PROGRAM MAIN
VAR

	fTotalCIP_Volume: REAL;
	fbWritePersistent: FB_WritePersistentData;
	bTesting		:	BOOL:=FALSE	;
	nI_1			: 	INT		;
	ftg_EStop_Fall	: 	F_TRIG	;
	rs_EStopFall	: 	RS	;
	bTestEstop		:	BOOL:=TRUE	;
	FB_OpenClose_Vlave_4026: FB_OpenClose_Vlave;
	bTemp_Water_Overweight_check: BOOL;
	fbUPS: FB_S_UPS_CX51x0;

	bSetExpeationTime: BOOL;
	i: E_ELEMENT_LIST;
	tExpirationSet_Test: TIME := T#10s;
END_VAR

prg_RealClock();
prg_Piston();
prg_Safety();
prg_MessageManager();
prg_Messages();
prg_Call_OpMode();
prg_IntCheck();
prg_User();
act_ResetPumps();
(*
prg_TriBlender(
		fb_TriBlenderPump:= g_Pump.fbPump[E_Pump_List.TB0001],
		stTriblender:=stTriblender,
		arrComponents:=arrProductionComponents);
*)		
//act_SetAnalogSens_Test();//To be deleted, for testing purposes
act_Call_Sensors_Analog();//To be deleted, for testing purposes
act_Call_Sensors_Analog_1();//To be deleted, for testing purposes
act_Call_ScaleFactor();//To be deleted, for testing purposes
act_Call_ProcessCntrl();

act_SetValves();
act_ClientPump_Select();
act_ClientStirrer_Select();
act_Call_Elements();
act_Call_Elements_Imp();
act_Call_Pumps();
prg_InterCon_Usage();
act_Sensors();
act_HeatExchenger();
act_Call_CIP();
act_Call_Production();

act_Call_For_HMI();

g_SFC.fbSFC_Temp1();

//Temtprary Overweght protection!!!!! DO NOT DELETE
IF fTotalCIP_Volume >=1500 AND FALSE THEN;
	//fbPis[E_Pis_Name.V1022].m_SetByRecipe(stPis:=stPis[E_Pis_Name.V1022], req:=E_Piston_Recipe_State.Release);
	//fbPis[E_Pis_Name.V1019].m_SetByRecipe(stPis:=stPis[E_Pis_Name.V1019], req:=E_Piston_Recipe_State.Release);
	//fbPis[E_Pis_Name.V1016].m_SetByRecipe(stPis:=stPis[E_Pis_Name.V1016], req:=E_Piston_Recipe_State.Release);
	//fbPis[E_Pis_Name.V1011].m_SetByRecipe(stPis:=stPis[E_Pis_Name.V1011], req:=E_Piston_Recipe_State.Release);
	bTemp_Water_Overweight_check:=FALSE;
	fbPrintErrMessageByID(sModuleDescription:='CIP',sActErrorID:='101x000x000');
ELSIF fTotalCIP_Volume < 1480 THEN;
	bTemp_Water_Overweight_check:=TRUE;
END_IF

IF arrTanksSens[E_Tank_Name.T91].get_stTankLevel_OverFlow() THEN;
	fbPis[E_Pis_Name.V1022].m_SetByRecipe(stPis:=stPis[E_Pis_Name.V1022], req:=E_Piston_Recipe_State.Release);
	//print error
	fbPrintErrMessageByID(sModuleDescription:='CIP',sActErrorID:='101x000x001');		
END_IF
IF arrTanksSens[E_Tank_Name.T92].get_stTankLevel_OverFlow() THEN;
	fbPis[E_Pis_Name.V1019].m_SetByRecipe(stPis:=stPis[E_Pis_Name.V1019], req:=E_Piston_Recipe_State.Release);
	//print error
	fbPrintErrMessageByID(sModuleDescription:='CIP',sActErrorID:='101x000x002');		
END_IF
IF arrTanksSens[E_Tank_Name.T93].get_stTankLevel_OverFlow() THEN;
	fbPis[E_Pis_Name.V1016].m_SetByRecipe(stPis:=stPis[E_Pis_Name.V1016], req:=E_Piston_Recipe_State.Release);
	//print error	
	fbPrintErrMessageByID(sModuleDescription:='CIP',sActErrorID:='101x000x003');	
END_IF
IF arrTanksSens[E_Tank_Name.T94].get_stTankLevel_OverFlow() THEN;
	fbPis[E_Pis_Name.V1011].m_SetByRecipe(stPis:=stPis[E_Pis_Name.V1011], req:=E_Piston_Recipe_State.Release);
	//print error
	fbPrintErrMessageByID(sModuleDescription:='CIP',sActErrorID:='101x000x004');		
END_IF
	
IF bSetExpeationTime THEN;
	bSetExpeationTime:=FALSE;
	FOR i:=E_Element_List.eTank_1 TO E_Element_List.eLine_Color DO
		fbElement[i].ExpirationTime:=tExpirationSet_Test;
		
	END_FOR
END_IF
	

mElementList_SetName();

fbWritePersistent(
	NETID:= , 
	PORT:= 851, 
	START:= , 
	TMOUT:= T#3S, 
	MODE:= , 
	BUSY=> , 
	ERR=> , 
	ERRID=> );

fbUPS();

ACTION act_Call_CIP:
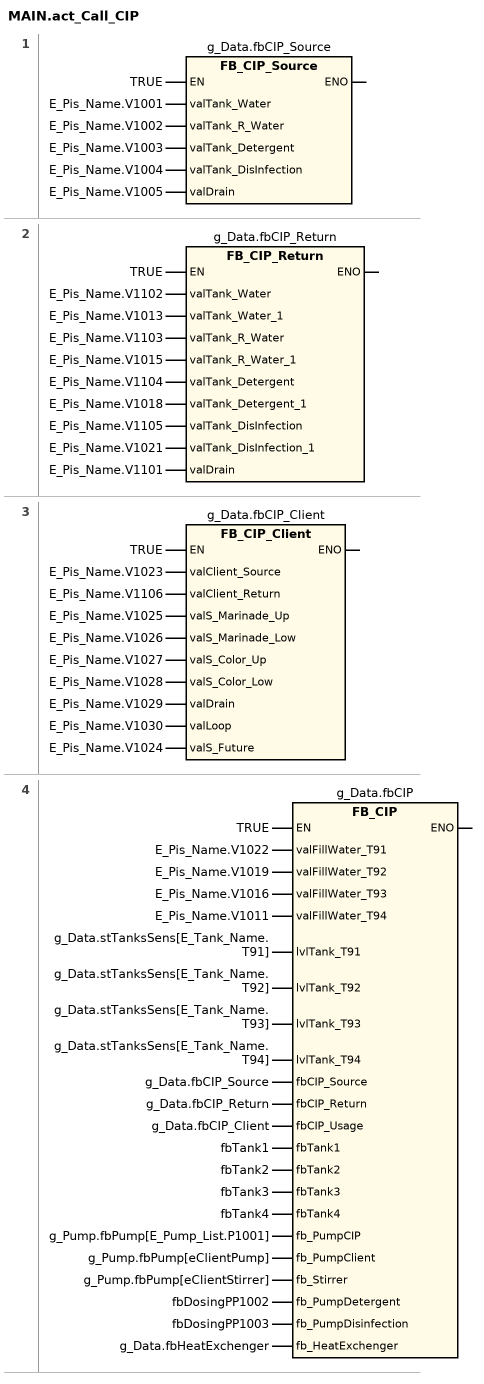
// NETWORK 1
g_Data.fbCIP_Source(
    valTank_Water := E_Pis_Name.V1001,
    valTank_R_Water := E_Pis_Name.V1002,
    valTank_Detergent := E_Pis_Name.V1003,
    valTank_DisInfection := E_Pis_Name.V1004,
    valDrain := E_Pis_Name.V1005); // FB_CIP_Source

// NETWORK 2
g_Data.fbCIP_Return(
    valTank_Water := E_Pis_Name.V1102,
    valTank_Water_1 := E_Pis_Name.V1013,
    valTank_R_Water := E_Pis_Name.V1103,
    valTank_R_Water_1 := E_Pis_Name.V1015,
    valTank_Detergent := E_Pis_Name.V1104,
    valTank_Detergent_1 := E_Pis_Name.V1018,
    valTank_DisInfection := E_Pis_Name.V1105,
    valTank_DisInfection_1 := E_Pis_Name.V1021,
    valDrain := E_Pis_Name.V1101); // FB_CIP_Return

// NETWORK 3
g_Data.fbCIP_Client(
    valClient_Source := E_Pis_Name.V1023,
    valClient_Return := E_Pis_Name.V1106,
    valS_Marinade_Up := E_Pis_Name.V1025,
    valS_Marinade_Low := E_Pis_Name.V1026,
    valS_Color_Up := E_Pis_Name.V1027,
    valS_Color_Low := E_Pis_Name.V1028,
    valDrain := E_Pis_Name.V1029,
    valLoop := E_Pis_Name.V1030,
    valS_Future := E_Pis_Name.V1024); // FB_CIP_Client

// NETWORK 4
g_Data.fbCIP(
    valFillWater_T91 := E_Pis_Name.V1022,
    valFillWater_T92 := E_Pis_Name.V1019,
    valFillWater_T93 := E_Pis_Name.V1016,
    valFillWater_T94 := E_Pis_Name.V1011,
    lvlTank_T91 := g_Data.stTanksSens[E_Tank_Name.T91],
    lvlTank_T92 := g_Data.stTanksSens[E_Tank_Name.T92],
    lvlTank_T93 := g_Data.stTanksSens[E_Tank_Name.T93],
    lvlTank_T94 := g_Data.stTanksSens[E_Tank_Name.T94],
    fbCIP_Source := g_Data.fbCIP_Source,
    fbCIP_Return := g_Data.fbCIP_Return,
    fbCIP_Usage := g_Data.fbCIP_Client,
    fbTank1 := fbTank1,
    fbTank2 := fbTank2,
    fbTank3 := fbTank3,
    fbTank4 := fbTank4,
    fb_PumpCIP := g_Pump.fbPump[E_Pump_List.P1001],
    fb_PumpClient := g_Pump.fbPump[eClientPump],
    fb_Stirrer := g_Pump.fbPump[eClientStirrer],
    fb_PumpDetergent := fbDosingPP1002,
    fb_PumpDisinfection := fbDosingPP1003,
    fb_HeatExchenger := g_Data.fbHeatExchenger); // FB_CIP

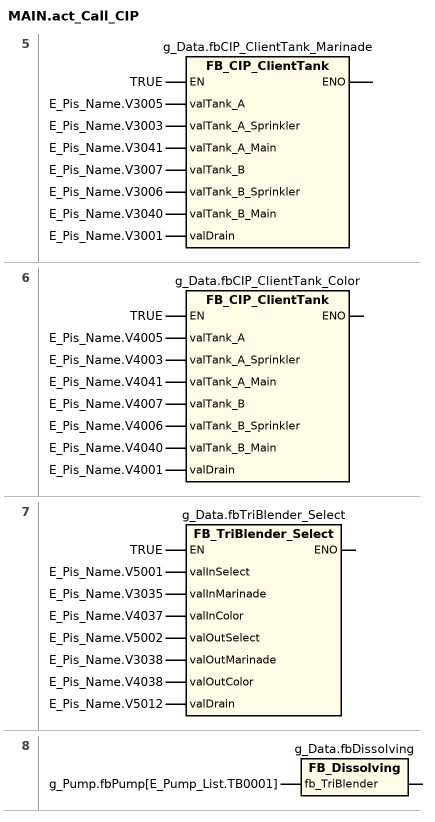
// NETWORK 5
g_Data.fbCIP_ClientTank_Marinade(
    valTank_A := E_Pis_Name.V3005,
    valTank_A_Sprinkler := E_Pis_Name.V3003,
    valTank_A_Main := E_Pis_Name.V3041,
    valTank_B := E_Pis_Name.V3007,
    valTank_B_Sprinkler := E_Pis_Name.V3006,
    valTank_B_Main := E_Pis_Name.V3040,
    valDrain := E_Pis_Name.V3001); // FB_CIP_ClientTank

// NETWORK 6
g_Data.fbCIP_ClientTank_Color(
    valTank_A := E_Pis_Name.V4005,
    valTank_A_Sprinkler := E_Pis_Name.V4003,
    valTank_A_Main := E_Pis_Name.V4041,
    valTank_B := E_Pis_Name.V4007,
    valTank_B_Sprinkler := E_Pis_Name.V4006,
    valTank_B_Main := E_Pis_Name.V4040,
    valDrain := E_Pis_Name.V4001); // FB_CIP_ClientTank

// NETWORK 7
g_Data.fbTriBlender_Select(
    valInSelect := E_Pis_Name.V5001,
    valInMarinade := E_Pis_Name.V3035,
    valInColor := E_Pis_Name.V4037,
    valOutSelect := E_Pis_Name.V5002,
    valOutMarinade := E_Pis_Name.V3038,
    valOutColor := E_Pis_Name.V4038,
    valDrain := E_Pis_Name.V5012); // FB_TriBlender_Select

// NETWORK 8
g_Data.fbDissolving(fb_TriBlender := g_Pump.fbPump[E_Pump_List.TB0001]); // FB_Dissolving
END_ACTION

ACTION act_Call_Elements:
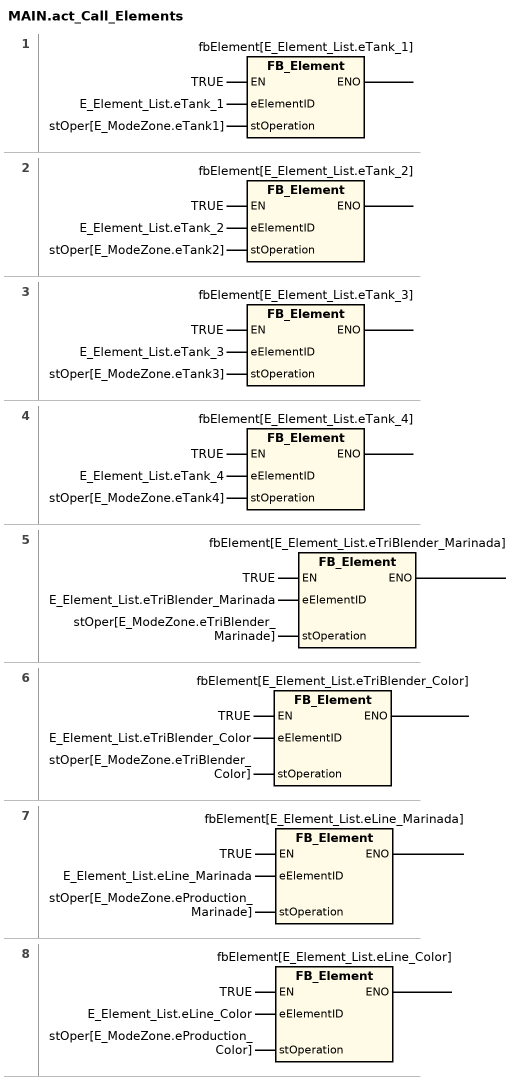
// NETWORK 1
fbElement[E_Element_List.eTank_1](eElementID := E_Element_List.eTank_1, stOperation := stOper[E_ModeZone.eTank1]); // FB_Element

// NETWORK 2
fbElement[E_Element_List.eTank_2](eElementID := E_Element_List.eTank_2, stOperation := stOper[E_ModeZone.eTank2]); // FB_Element

// NETWORK 3
fbElement[E_Element_List.eTank_3](eElementID := E_Element_List.eTank_3, stOperation := stOper[E_ModeZone.eTank3]); // FB_Element

// NETWORK 4
fbElement[E_Element_List.eTank_4](eElementID := E_Element_List.eTank_4, stOperation := stOper[E_ModeZone.eTank4]); // FB_Element

// NETWORK 5
fbElement[E_Element_List.eTriBlender_Marinada](eElementID := E_Element_List.eTriBlender_Marinada, stOperation := stOper[E_ModeZone.eTriBlender_Marinade]); // FB_Element

// NETWORK 6
fbElement[E_Element_List.eTriBlender_Color](eElementID := E_Element_List.eTriBlender_Color, stOperation := stOper[E_ModeZone.eTriBlender_Color]); // FB_Element

// NETWORK 7
fbElement[E_Element_List.eLine_Marinada](eElementID := E_Element_List.eLine_Marinada, stOperation := stOper[E_ModeZone.eProduction_Marinade]); // FB_Element

// NETWORK 8
fbElement[E_Element_List.eLine_Color](eElementID := E_Element_List.eLine_Color, stOperation := stOper[E_ModeZone.eProduction_Color]); // FB_Element
END_ACTION

ACTION act_Call_Elements_Imp:
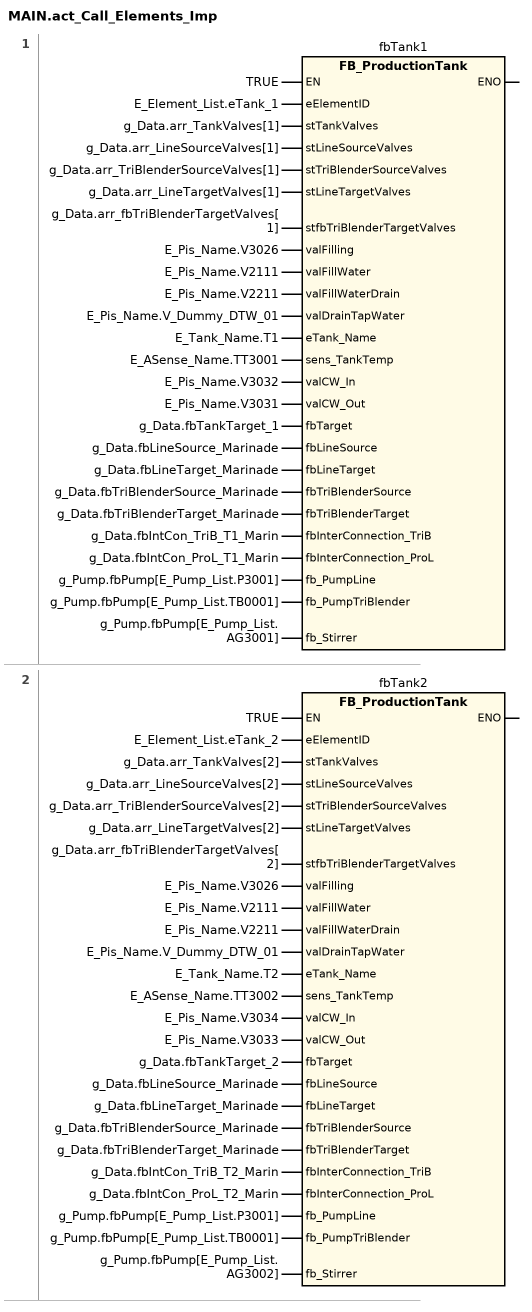
// NETWORK 1
fbTank1(
    eElementID := E_Element_List.eTank_1,
    stTankValves := g_Data.arr_TankValves[1],
    stLineSourceValves := g_Data.arr_LineSourceValves[1],
    stTriBlenderSourceValves := g_Data.arr_TriBlenderSourceValves[1],
    stLineTargetValves := g_Data.arr_LineTargetValves[1],
    stfbTriBlenderTargetValves := g_Data.arr_fbTriBlenderTargetValves[1],
    valFilling := E_Pis_Name.V3026,
    valFillWater := E_Pis_Name.V2111,
    valFillWaterDrain := E_Pis_Name.V2211,
    valDrainTapWater := E_Pis_Name.V_Dummy_DTW_01,
    eTank_Name := E_Tank_Name.T1,
    sens_TankTemp := E_ASense_Name.TT3001,
    valCW_In := E_Pis_Name.V3032,
    valCW_Out := E_Pis_Name.V3031,
    fbTarget := g_Data.fbTankTarget_1,
    fbLineSource := g_Data.fbLineSource_Marinade,
    fbLineTarget := g_Data.fbLineTarget_Marinade,
    fbTriBlenderSource := g_Data.fbTriBlenderSource_Marinade,
    fbTriBlenderTarget := g_Data.fbTriBlenderTarget_Marinade,
    fbInterConnection_TriB := g_Data.fbIntCon_TriB_T1_Marin,
    fbInterConnection_ProL := g_Data.fbIntCon_ProL_T1_Marin,
    fb_PumpLine := g_Pump.fbPump[E_Pump_List.P3001],
    fb_PumpTriBlender := g_Pump.fbPump[E_Pump_List.TB0001],
    fb_Stirrer := g_Pump.fbPump[E_Pump_List.AG3001]); // FB_ProductionTank

// NETWORK 2
fbTank2(
    eElementID := E_Element_List.eTank_2,
    stTankValves := g_Data.arr_TankValves[2],
    stLineSourceValves := g_Data.arr_LineSourceValves[2],
    stTriBlenderSourceValves := g_Data.arr_TriBlenderSourceValves[2],
    stLineTargetValves := g_Data.arr_LineTargetValves[2],
    stfbTriBlenderTargetValves := g_Data.arr_fbTriBlenderTargetValves[2],
    valFilling := E_Pis_Name.V3026,
    valFillWater := E_Pis_Name.V2111,
    valFillWaterDrain := E_Pis_Name.V2211,
    valDrainTapWater := E_Pis_Name.V_Dummy_DTW_01,
    eTank_Name := E_Tank_Name.T2,
    sens_TankTemp := E_ASense_Name.TT3002,
    valCW_In := E_Pis_Name.V3034,
    valCW_Out := E_Pis_Name.V3033,
    fbTarget := g_Data.fbTankTarget_2,
    fbLineSource := g_Data.fbLineSource_Marinade,
    fbLineTarget := g_Data.fbLineTarget_Marinade,
    fbTriBlenderSource := g_Data.fbTriBlenderSource_Marinade,
    fbTriBlenderTarget := g_Data.fbTriBlenderTarget_Marinade,
    fbInterConnection_TriB := g_Data.fbIntCon_TriB_T2_Marin,
    fbInterConnection_ProL := g_Data.fbIntCon_ProL_T2_Marin,
    fb_PumpLine := g_Pump.fbPump[E_Pump_List.P3001],
    fb_PumpTriBlender := g_Pump.fbPump[E_Pump_List.TB0001],
    fb_Stirrer := g_Pump.fbPump[E_Pump_List.AG3002]); // FB_ProductionTank

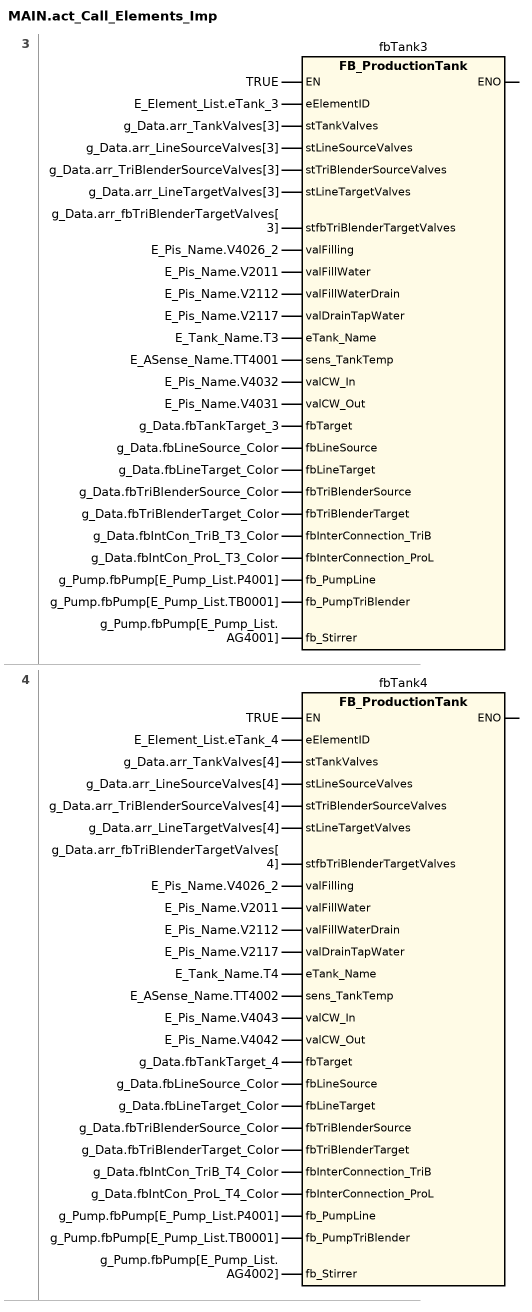
// NETWORK 3
fbTank3(
    eElementID := E_Element_List.eTank_3,
    stTankValves := g_Data.arr_TankValves[3],
    stLineSourceValves := g_Data.arr_LineSourceValves[3],
    stTriBlenderSourceValves := g_Data.arr_TriBlenderSourceValves[3],
    stLineTargetValves := g_Data.arr_LineTargetValves[3],
    stfbTriBlenderTargetValves := g_Data.arr_fbTriBlenderTargetValves[3],
    valFilling := E_Pis_Name.V4026_2,
    valFillWater := E_Pis_Name.V2011,
    valFillWaterDrain := E_Pis_Name.V2112,
    valDrainTapWater := E_Pis_Name.V2117,
    eTank_Name := E_Tank_Name.T3,
    sens_TankTemp := E_ASense_Name.TT4001,
    valCW_In := E_Pis_Name.V4032,
    valCW_Out := E_Pis_Name.V4031,
    fbTarget := g_Data.fbTankTarget_3,
    fbLineSource := g_Data.fbLineSource_Color,
    fbLineTarget := g_Data.fbLineTarget_Color,
    fbTriBlenderSource := g_Data.fbTriBlenderSource_Color,
    fbTriBlenderTarget := g_Data.fbTriBlenderTarget_Color,
    fbInterConnection_TriB := g_Data.fbIntCon_TriB_T3_Color,
    fbInterConnection_ProL := g_Data.fbIntCon_ProL_T3_Color,
    fb_PumpLine := g_Pump.fbPump[E_Pump_List.P4001],
    fb_PumpTriBlender := g_Pump.fbPump[E_Pump_List.TB0001],
    fb_Stirrer := g_Pump.fbPump[E_Pump_List.AG4001]); // FB_ProductionTank

// NETWORK 4
fbTank4(
    eElementID := E_Element_List.eTank_4,
    stTankValves := g_Data.arr_TankValves[4],
    stLineSourceValves := g_Data.arr_LineSourceValves[4],
    stTriBlenderSourceValves := g_Data.arr_TriBlenderSourceValves[4],
    stLineTargetValves := g_Data.arr_LineTargetValves[4],
    stfbTriBlenderTargetValves := g_Data.arr_fbTriBlenderTargetValves[4],
    valFilling := E_Pis_Name.V4026_2,
    valFillWater := E_Pis_Name.V2011,
    valFillWaterDrain := E_Pis_Name.V2112,
    valDrainTapWater := E_Pis_Name.V2117,
    eTank_Name := E_Tank_Name.T4,
    sens_TankTemp := E_ASense_Name.TT4002,
    valCW_In := E_Pis_Name.V4043,
    valCW_Out := E_Pis_Name.V4042,
    fbTarget := g_Data.fbTankTarget_4,
    fbLineSource := g_Data.fbLineSource_Color,
    fbLineTarget := g_Data.fbLineTarget_Color,
    fbTriBlenderSource := g_Data.fbTriBlenderSource_Color,
    fbTriBlenderTarget := g_Data.fbTriBlenderTarget_Color,
    fbInterConnection_TriB := g_Data.fbIntCon_TriB_T4_Color,
    fbInterConnection_ProL := g_Data.fbIntCon_ProL_T4_Color,
    fb_PumpLine := g_Pump.fbPump[E_Pump_List.P4001],
    fb_PumpTriBlender := g_Pump.fbPump[E_Pump_List.TB0001],
    fb_Stirrer := g_Pump.fbPump[E_Pump_List.AG4002]); // FB_ProductionTank
END_ACTION

ACTION act_Call_For_HMI:


g_HMI.stT91_Sens:=g_Data.stTanksSens[E_Tank_Name.T91];
g_HMI.stT92_Sens:=g_Data.stTanksSens[E_Tank_Name.T92];
g_HMI.stT93_Sens:=g_Data.stTanksSens[E_Tank_Name.T93];
g_HMI.stT94_Sens:=g_Data.stTanksSens[E_Tank_Name.T94];

g_HMI.stT1_Sens:=g_Data.stTanksSens[E_Tank_Name.T1];
g_HMI.stT2_Sens:=g_Data.stTanksSens[E_Tank_Name.T2];
g_HMI.stT3_Sens:=g_Data.stTanksSens[E_Tank_Name.T3];
g_HMI.stT4_Sens:=g_Data.stTanksSens[E_Tank_Name.T4];
END_ACTION

ACTION act_Call_ProcessCntrl:
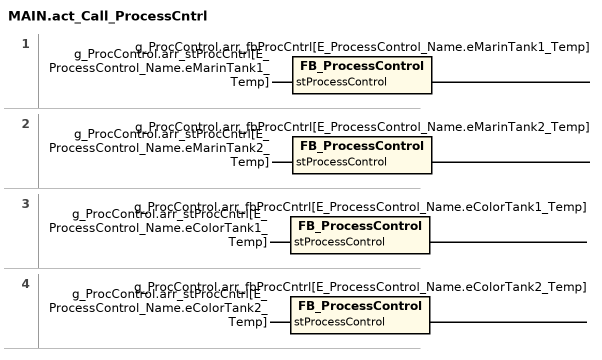
// NETWORK 1
g_ProcControl.arr_fbProcCntrl[E_ProcessControl_Name.eMarinTank1_Temp](stProcessControl := g_ProcControl.arr_stProcCntrl[E_ProcessControl_Name.eMarinTank1_Temp]); // FB_ProcessControl

// NETWORK 2
g_ProcControl.arr_fbProcCntrl[E_ProcessControl_Name.eMarinTank2_Temp](stProcessControl := g_ProcControl.arr_stProcCntrl[E_ProcessControl_Name.eMarinTank2_Temp]); // FB_ProcessControl

// NETWORK 3
g_ProcControl.arr_fbProcCntrl[E_ProcessControl_Name.eColorTank1_Temp](stProcessControl := g_ProcControl.arr_stProcCntrl[E_ProcessControl_Name.eColorTank1_Temp]); // FB_ProcessControl

// NETWORK 4
g_ProcControl.arr_fbProcCntrl[E_ProcessControl_Name.eColorTank2_Temp](stProcessControl := g_ProcControl.arr_stProcCntrl[E_ProcessControl_Name.eColorTank2_Temp]); // FB_ProcessControl
END_ACTION

ACTION act_Call_Production:

g_Prod.fbProdRecipe_Manage();
END_ACTION

ACTION act_Call_Pump_TB:
IF fbElement[E_Element_List.eTriBlender_Color].m_Get_InterConnection()=E_InterConnection.ConnToCIP 
OR fbElement[E_Element_List.eTriBlender_Marinada].m_Get_InterConnection()=E_InterConnection.ConnToCIP 
OR FALSE
THEN;
	act_Call_Pump_TB_CIP();
ELSE;
	CASE g_Data.eTriBlenderUsage OF
		E_TriBlenderUsage.eMarinada_T1,E_TriBlenderUsage.eMarinada_T2:;
				act_Call_Pump_TB_M();
		E_TriBlenderUsage.eColor_T3,E_TriBlenderUsage.eColor_T4:;
				act_Call_Pump_TB_C();
	ELSE;
		act_Call_Pump_TB_0();
	END_CASE	
END_IF
END_ACTION

ACTION act_Call_Pump_TB_0:
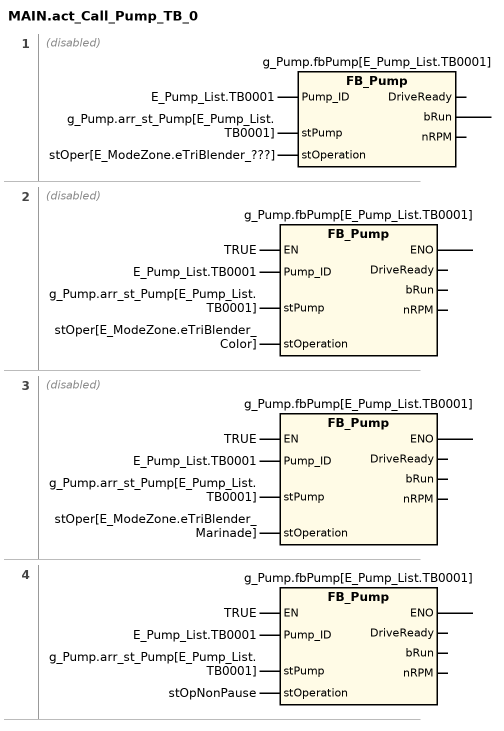
// NETWORK 1 (disabled)
// g_Pump.fbPump[E_Pump_List.TB0001](
//     Pump_ID := E_Pump_List.TB0001,
//     stPump := g_Pump.arr_st_Pump[E_Pump_List.TB0001],
//     stOperation := stOper[E_ModeZone.eTriBlender_???]); // FB_Pump

// NETWORK 2 (disabled)
// g_Pump.fbPump[E_Pump_List.TB0001](
//     Pump_ID := E_Pump_List.TB0001,
//     stPump := g_Pump.arr_st_Pump[E_Pump_List.TB0001],
//     stOperation := stOper[E_ModeZone.eTriBlender_Color]); // FB_Pump

// NETWORK 3 (disabled)
// g_Pump.fbPump[E_Pump_List.TB0001](
//     Pump_ID := E_Pump_List.TB0001,
//     stPump := g_Pump.arr_st_Pump[E_Pump_List.TB0001],
//     stOperation := stOper[E_ModeZone.eTriBlender_Marinade]); // FB_Pump

// NETWORK 4
g_Pump.fbPump[E_Pump_List.TB0001](
    Pump_ID := E_Pump_List.TB0001,
    stPump := g_Pump.arr_st_Pump[E_Pump_List.TB0001],
    stOperation := stOpNonPause); // FB_Pump
END_ACTION

ACTION act_Call_Pump_TB_C:
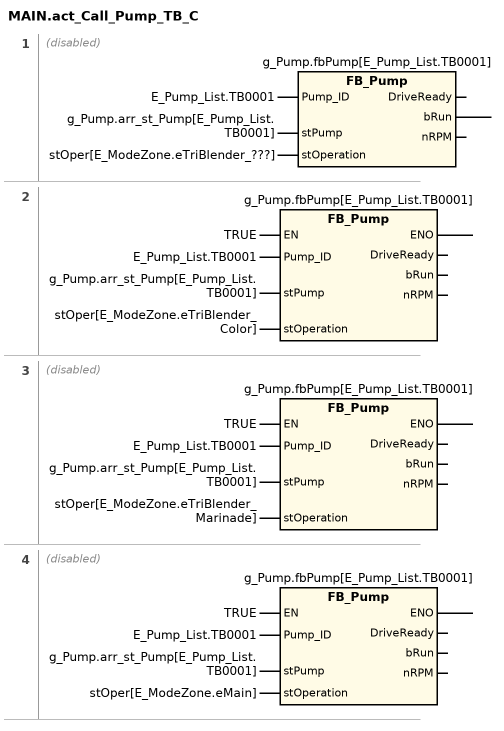
// NETWORK 1 (disabled)
// g_Pump.fbPump[E_Pump_List.TB0001](
//     Pump_ID := E_Pump_List.TB0001,
//     stPump := g_Pump.arr_st_Pump[E_Pump_List.TB0001],
//     stOperation := stOper[E_ModeZone.eTriBlender_???]); // FB_Pump

// NETWORK 2
g_Pump.fbPump[E_Pump_List.TB0001](
    Pump_ID := E_Pump_List.TB0001,
    stPump := g_Pump.arr_st_Pump[E_Pump_List.TB0001],
    stOperation := stOper[E_ModeZone.eTriBlender_Color]); // FB_Pump

// NETWORK 3 (disabled)
// g_Pump.fbPump[E_Pump_List.TB0001](
//     Pump_ID := E_Pump_List.TB0001,
//     stPump := g_Pump.arr_st_Pump[E_Pump_List.TB0001],
//     stOperation := stOper[E_ModeZone.eTriBlender_Marinade]); // FB_Pump

// NETWORK 4 (disabled)
// g_Pump.fbPump[E_Pump_List.TB0001](
//     Pump_ID := E_Pump_List.TB0001,
//     stPump := g_Pump.arr_st_Pump[E_Pump_List.TB0001],
//     stOperation := stOper[E_ModeZone.eMain]); // FB_Pump
END_ACTION

ACTION act_Call_Pump_TB_CIP:
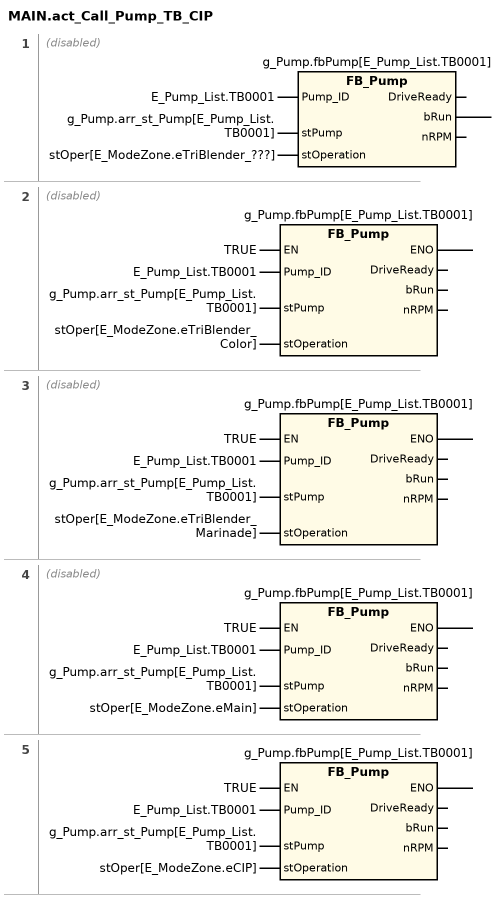
// NETWORK 1 (disabled)
// g_Pump.fbPump[E_Pump_List.TB0001](
//     Pump_ID := E_Pump_List.TB0001,
//     stPump := g_Pump.arr_st_Pump[E_Pump_List.TB0001],
//     stOperation := stOper[E_ModeZone.eTriBlender_???]); // FB_Pump

// NETWORK 2 (disabled)
// g_Pump.fbPump[E_Pump_List.TB0001](
//     Pump_ID := E_Pump_List.TB0001,
//     stPump := g_Pump.arr_st_Pump[E_Pump_List.TB0001],
//     stOperation := stOper[E_ModeZone.eTriBlender_Color]); // FB_Pump

// NETWORK 3 (disabled)
// g_Pump.fbPump[E_Pump_List.TB0001](
//     Pump_ID := E_Pump_List.TB0001,
//     stPump := g_Pump.arr_st_Pump[E_Pump_List.TB0001],
//     stOperation := stOper[E_ModeZone.eTriBlender_Marinade]); // FB_Pump

// NETWORK 4 (disabled)
// g_Pump.fbPump[E_Pump_List.TB0001](
//     Pump_ID := E_Pump_List.TB0001,
//     stPump := g_Pump.arr_st_Pump[E_Pump_List.TB0001],
//     stOperation := stOper[E_ModeZone.eMain]); // FB_Pump

// NETWORK 5
g_Pump.fbPump[E_Pump_List.TB0001](
    Pump_ID := E_Pump_List.TB0001,
    stPump := g_Pump.arr_st_Pump[E_Pump_List.TB0001],
    stOperation := stOper[E_ModeZone.eCIP]); // FB_Pump
END_ACTION

ACTION act_Call_Pump_TB_M:
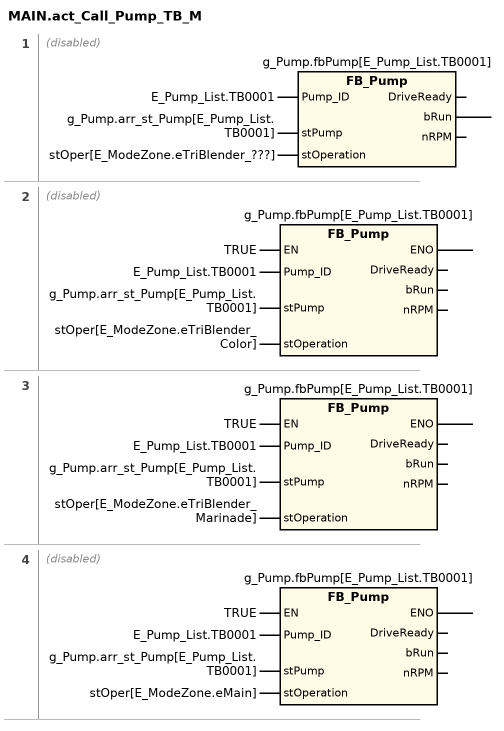
// NETWORK 1 (disabled)
// g_Pump.fbPump[E_Pump_List.TB0001](
//     Pump_ID := E_Pump_List.TB0001,
//     stPump := g_Pump.arr_st_Pump[E_Pump_List.TB0001],
//     stOperation := stOper[E_ModeZone.eTriBlender_???]); // FB_Pump

// NETWORK 2 (disabled)
// g_Pump.fbPump[E_Pump_List.TB0001](
//     Pump_ID := E_Pump_List.TB0001,
//     stPump := g_Pump.arr_st_Pump[E_Pump_List.TB0001],
//     stOperation := stOper[E_ModeZone.eTriBlender_Color]); // FB_Pump

// NETWORK 3
g_Pump.fbPump[E_Pump_List.TB0001](
    Pump_ID := E_Pump_List.TB0001,
    stPump := g_Pump.arr_st_Pump[E_Pump_List.TB0001],
    stOperation := stOper[E_ModeZone.eTriBlender_Marinade]); // FB_Pump

// NETWORK 4 (disabled)
// g_Pump.fbPump[E_Pump_List.TB0001](
//     Pump_ID := E_Pump_List.TB0001,
//     stPump := g_Pump.arr_st_Pump[E_Pump_List.TB0001],
//     stOperation := stOper[E_ModeZone.eMain]); // FB_Pump
END_ACTION

ACTION act_Call_Pumps:
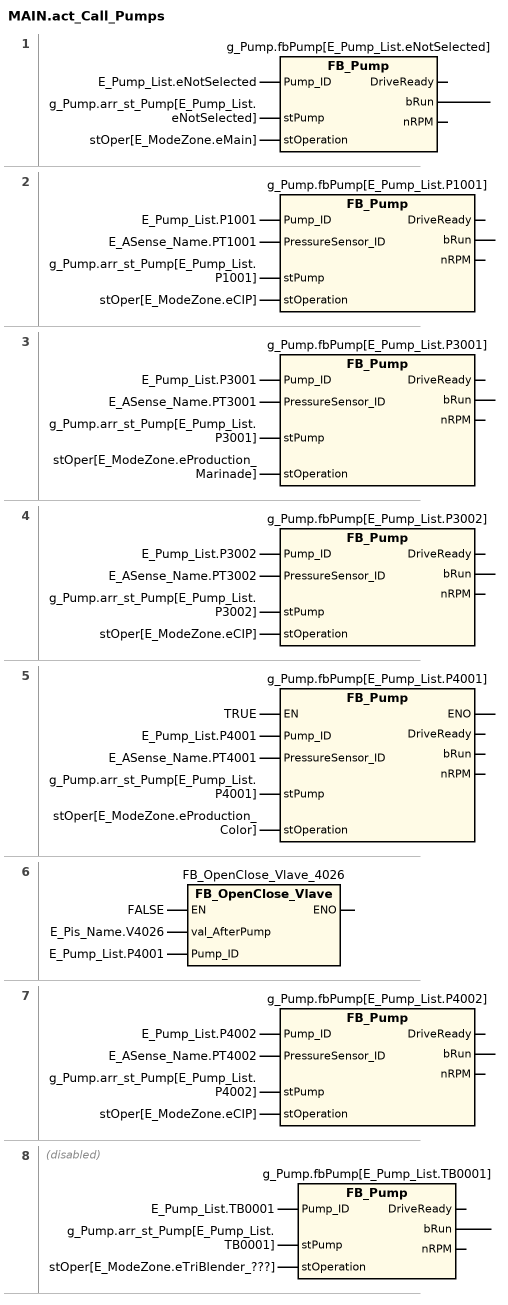
// NETWORK 1
g_Pump.fbPump[E_Pump_List.eNotSelected](
    Pump_ID := E_Pump_List.eNotSelected,
    stPump := g_Pump.arr_st_Pump[E_Pump_List.eNotSelected],
    stOperation := stOper[E_ModeZone.eMain]); // FB_Pump

// NETWORK 2
g_Pump.fbPump[E_Pump_List.P1001](
    Pump_ID := E_Pump_List.P1001,
    PressureSensor_ID := E_ASense_Name.PT1001,
    stPump := g_Pump.arr_st_Pump[E_Pump_List.P1001],
    stOperation := stOper[E_ModeZone.eCIP]); // FB_Pump

// NETWORK 3
g_Pump.fbPump[E_Pump_List.P3001](
    Pump_ID := E_Pump_List.P3001,
    PressureSensor_ID := E_ASense_Name.PT3001,
    stPump := g_Pump.arr_st_Pump[E_Pump_List.P3001],
    stOperation := stOper[E_ModeZone.eProduction_Marinade]); // FB_Pump

// NETWORK 4
g_Pump.fbPump[E_Pump_List.P3002](
    Pump_ID := E_Pump_List.P3002,
    PressureSensor_ID := E_ASense_Name.PT3002,
    stPump := g_Pump.arr_st_Pump[E_Pump_List.P3002],
    stOperation := stOper[E_ModeZone.eCIP]); // FB_Pump

// NETWORK 5
g_Pump.fbPump[E_Pump_List.P4001](
    Pump_ID := E_Pump_List.P4001,
    PressureSensor_ID := E_ASense_Name.PT4001,
    stPump := g_Pump.arr_st_Pump[E_Pump_List.P4001],
    stOperation := stOper[E_ModeZone.eProduction_Color]); // FB_Pump

// NETWORK 6
IF FALSE THEN
    FB_OpenClose_Vlave_4026(val_AfterPump := E_Pis_Name.V4026, Pump_ID := E_Pump_List.P4001); // FB_OpenClose_Vlave
END_IF

// NETWORK 7
g_Pump.fbPump[E_Pump_List.P4002](
    Pump_ID := E_Pump_List.P4002,
    PressureSensor_ID := E_ASense_Name.PT4002,
    stPump := g_Pump.arr_st_Pump[E_Pump_List.P4002],
    stOperation := stOper[E_ModeZone.eCIP]); // FB_Pump

// NETWORK 8 (disabled)
// g_Pump.fbPump[E_Pump_List.TB0001](
//     Pump_ID := E_Pump_List.TB0001,
//     stPump := g_Pump.arr_st_Pump[E_Pump_List.TB0001],
//     stOperation := stOper[E_ModeZone.eTriBlender_???]); // FB_Pump

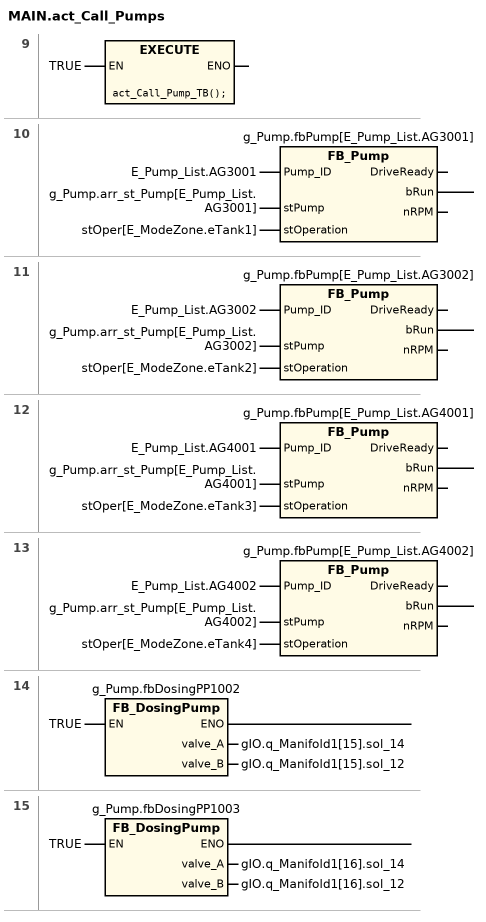
// NETWORK 9

act_Call_Pump_TB();

// NETWORK 10
g_Pump.fbPump[E_Pump_List.AG3001](
    Pump_ID := E_Pump_List.AG3001,
    stPump := g_Pump.arr_st_Pump[E_Pump_List.AG3001],
    stOperation := stOper[E_ModeZone.eTank1]); // FB_Pump

// NETWORK 11
g_Pump.fbPump[E_Pump_List.AG3002](
    Pump_ID := E_Pump_List.AG3002,
    stPump := g_Pump.arr_st_Pump[E_Pump_List.AG3002],
    stOperation := stOper[E_ModeZone.eTank2]); // FB_Pump

// NETWORK 12
g_Pump.fbPump[E_Pump_List.AG4001](
    Pump_ID := E_Pump_List.AG4001,
    stPump := g_Pump.arr_st_Pump[E_Pump_List.AG4001],
    stOperation := stOper[E_ModeZone.eTank3]); // FB_Pump

// NETWORK 13
g_Pump.fbPump[E_Pump_List.AG4002](
    Pump_ID := E_Pump_List.AG4002,
    stPump := g_Pump.arr_st_Pump[E_Pump_List.AG4002],
    stOperation := stOper[E_ModeZone.eTank4]); // FB_Pump

// NETWORK 14
g_Pump.fbDosingPP1002(valve_A => gIO.q_Manifold1[15].sol_14, valve_B => gIO.q_Manifold1[15].sol_12); // FB_DosingPump

// NETWORK 15
g_Pump.fbDosingPP1003(valve_A => gIO.q_Manifold1[16].sol_14, valve_B => gIO.q_Manifold1[16].sol_12); // FB_DosingPump
END_ACTION

ACTION act_Call_ScaleFactor:
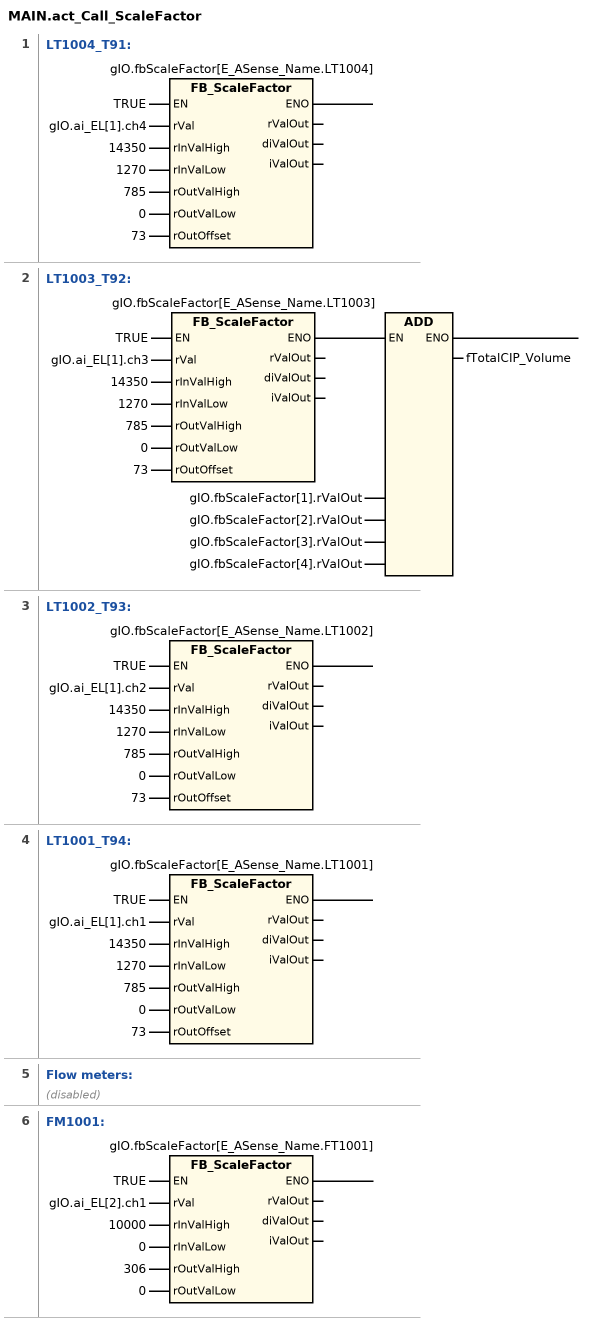
// NETWORK 1
LT1004_T91:
gIO.fbScaleFactor[E_ASense_Name.LT1004](
    rVal := gIO.ai_EL[1].ch4,
    rInValHigh := 14350,
    rInValLow := 1270,
    rOutValHigh := 785,
    rOutValLow := 0,
    rOutOffset := 73); // FB_ScaleFactor

// NETWORK 2
LT1003_T92:
gIO.fbScaleFactor[E_ASense_Name.LT1003](
    rVal := gIO.ai_EL[1].ch3,
    rInValHigh := 14350,
    rInValLow := 1270,
    rOutValHigh := 785,
    rOutValLow := 0,
    rOutOffset := 73); // FB_ScaleFactor
fTotalCIP_Volume := gIO.fbScaleFactor[1].rValOut + gIO.fbScaleFactor[2].rValOut + gIO.fbScaleFactor[3].rValOut + gIO.fbScaleFactor[4].rValOut;

// NETWORK 3
LT1002_T93:
gIO.fbScaleFactor[E_ASense_Name.LT1002](
    rVal := gIO.ai_EL[1].ch2,
    rInValHigh := 14350,
    rInValLow := 1270,
    rOutValHigh := 785,
    rOutValLow := 0,
    rOutOffset := 73); // FB_ScaleFactor

// NETWORK 4
LT1001_T94:
gIO.fbScaleFactor[E_ASense_Name.LT1001](
    rVal := gIO.ai_EL[1].ch1,
    rInValHigh := 14350,
    rInValLow := 1270,
    rOutValHigh := 785,
    rOutValLow := 0,
    rOutOffset := 73); // FB_ScaleFactor

// NETWORK 5 (disabled)
// label: Flow meters

// NETWORK 6
FM1001:
gIO.fbScaleFactor[E_ASense_Name.FT1001](
    rVal := gIO.ai_EL[2].ch1,
    rInValHigh := 10000,
    rInValLow := 0,
    rOutValHigh := 306,
    rOutValLow := 0); // FB_ScaleFactor

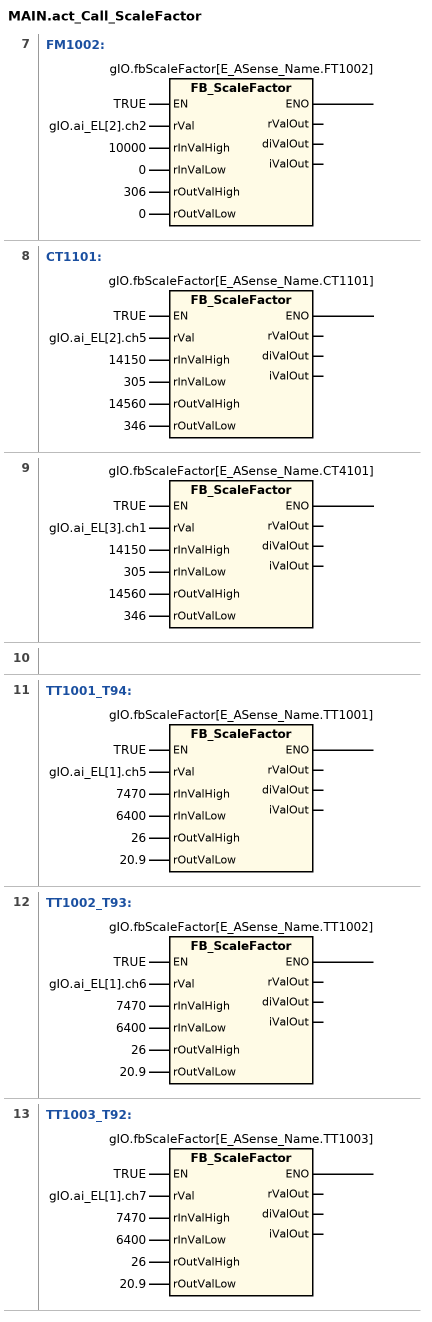
// NETWORK 7
FM1002:
gIO.fbScaleFactor[E_ASense_Name.FT1002](
    rVal := gIO.ai_EL[2].ch2,
    rInValHigh := 10000,
    rInValLow := 0,
    rOutValHigh := 306,
    rOutValLow := 0); // FB_ScaleFactor

// NETWORK 8
CT1101:
gIO.fbScaleFactor[E_ASense_Name.CT1101](
    rVal := gIO.ai_EL[2].ch5,
    rInValHigh := 14150,
    rInValLow := 305,
    rOutValHigh := 14560,
    rOutValLow := 346); // FB_ScaleFactor

// NETWORK 9
gIO.fbScaleFactor[E_ASense_Name.CT4101](
    rVal := gIO.ai_EL[3].ch1,
    rInValHigh := 14150,
    rInValLow := 305,
    rOutValHigh := 14560,
    rOutValLow := 346); // FB_ScaleFactor

// NETWORK 10

// NETWORK 11
TT1001_T94:
gIO.fbScaleFactor[E_ASense_Name.TT1001](
    rVal := gIO.ai_EL[1].ch5,
    rInValHigh := 7470,
    rInValLow := 6400,
    rOutValHigh := 26,
    rOutValLow := 20.9); // FB_ScaleFactor

// NETWORK 12
TT1002_T93:
gIO.fbScaleFactor[E_ASense_Name.TT1002](
    rVal := gIO.ai_EL[1].ch6,
    rInValHigh := 7470,
    rInValLow := 6400,
    rOutValHigh := 26,
    rOutValLow := 20.9); // FB_ScaleFactor

// NETWORK 13
TT1003_T92:
gIO.fbScaleFactor[E_ASense_Name.TT1003](
    rVal := gIO.ai_EL[1].ch7,
    rInValHigh := 7470,
    rInValLow := 6400,
    rOutValHigh := 26,
    rOutValLow := 20.9); // FB_ScaleFactor

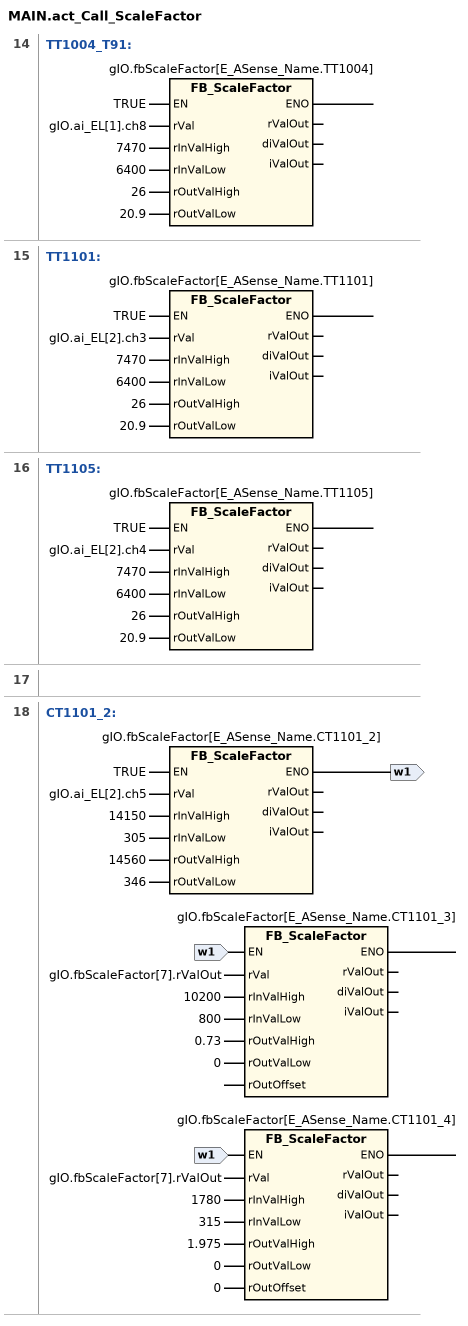
// NETWORK 14
TT1004_T91:
gIO.fbScaleFactor[E_ASense_Name.TT1004](
    rVal := gIO.ai_EL[1].ch8,
    rInValHigh := 7470,
    rInValLow := 6400,
    rOutValHigh := 26,
    rOutValLow := 20.9); // FB_ScaleFactor

// NETWORK 15
TT1101:
gIO.fbScaleFactor[E_ASense_Name.TT1101](
    rVal := gIO.ai_EL[2].ch3,
    rInValHigh := 7470,
    rInValLow := 6400,
    rOutValHigh := 26,
    rOutValLow := 20.9); // FB_ScaleFactor

// NETWORK 16
TT1105:
gIO.fbScaleFactor[E_ASense_Name.TT1105](
    rVal := gIO.ai_EL[2].ch4,
    rInValHigh := 7470,
    rInValLow := 6400,
    rOutValHigh := 26,
    rOutValLow := 20.9); // FB_ScaleFactor

// NETWORK 17

// NETWORK 18
CT1101_2:
gIO.fbScaleFactor[E_ASense_Name.CT1101_2](
    rVal := gIO.ai_EL[2].ch5,
    rInValHigh := 14150,
    rInValLow := 305,
    rOutValHigh := 14560,
    rOutValLow := 346); // FB_ScaleFactor
gIO.fbScaleFactor[E_ASense_Name.CT1101_3](
    rVal := gIO.fbScaleFactor[7].rValOut,
    rInValHigh := 10200,
    rInValLow := 800,
    rOutValHigh := 0.73,
    rOutValLow := 0); // FB_ScaleFactor
gIO.fbScaleFactor[E_ASense_Name.CT1101_4](
    rVal := gIO.fbScaleFactor[7].rValOut,
    rInValHigh := 1780,
    rInValLow := 315,
    rOutValHigh := 1.975,
    rOutValLow := 0,
    rOutOffset := 0); // FB_ScaleFactor

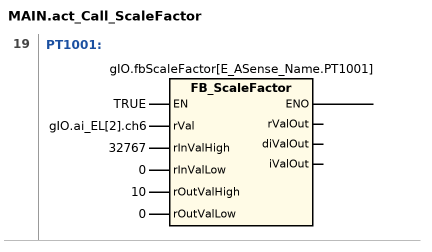
// NETWORK 19
PT1001:
gIO.fbScaleFactor[E_ASense_Name.PT1001](
    rVal := gIO.ai_EL[2].ch6,
    rInValHigh := 32767,
    rInValLow := 0,
    rOutValHigh := 10,
    rOutValLow := 0); // FB_ScaleFactor
END_ACTION

ACTION act_Call_Sensors_Analog:
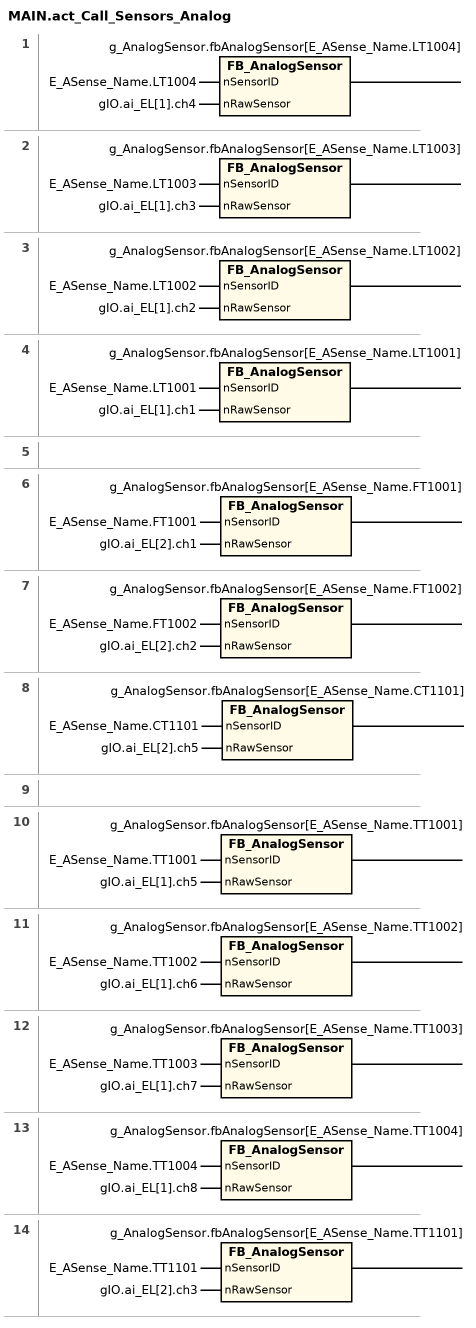
// NETWORK 1
g_AnalogSensor.fbAnalogSensor[E_ASense_Name.LT1004](nSensorID := E_ASense_Name.LT1004, nRawSensor := gIO.ai_EL[1].ch4); // FB_AnalogSensor

// NETWORK 2
g_AnalogSensor.fbAnalogSensor[E_ASense_Name.LT1003](nSensorID := E_ASense_Name.LT1003, nRawSensor := gIO.ai_EL[1].ch3); // FB_AnalogSensor

// NETWORK 3
g_AnalogSensor.fbAnalogSensor[E_ASense_Name.LT1002](nSensorID := E_ASense_Name.LT1002, nRawSensor := gIO.ai_EL[1].ch2); // FB_AnalogSensor

// NETWORK 4
g_AnalogSensor.fbAnalogSensor[E_ASense_Name.LT1001](nSensorID := E_ASense_Name.LT1001, nRawSensor := gIO.ai_EL[1].ch1); // FB_AnalogSensor

// NETWORK 5

// NETWORK 6
g_AnalogSensor.fbAnalogSensor[E_ASense_Name.FT1001](nSensorID := E_ASense_Name.FT1001, nRawSensor := gIO.ai_EL[2].ch1); // FB_AnalogSensor

// NETWORK 7
g_AnalogSensor.fbAnalogSensor[E_ASense_Name.FT1002](nSensorID := E_ASense_Name.FT1002, nRawSensor := gIO.ai_EL[2].ch2); // FB_AnalogSensor

// NETWORK 8
g_AnalogSensor.fbAnalogSensor[E_ASense_Name.CT1101](nSensorID := E_ASense_Name.CT1101, nRawSensor := gIO.ai_EL[2].ch5); // FB_AnalogSensor

// NETWORK 9

// NETWORK 10
g_AnalogSensor.fbAnalogSensor[E_ASense_Name.TT1001](nSensorID := E_ASense_Name.TT1001, nRawSensor := gIO.ai_EL[1].ch5); // FB_AnalogSensor

// NETWORK 11
g_AnalogSensor.fbAnalogSensor[E_ASense_Name.TT1002](nSensorID := E_ASense_Name.TT1002, nRawSensor := gIO.ai_EL[1].ch6); // FB_AnalogSensor

// NETWORK 12
g_AnalogSensor.fbAnalogSensor[E_ASense_Name.TT1003](nSensorID := E_ASense_Name.TT1003, nRawSensor := gIO.ai_EL[1].ch7); // FB_AnalogSensor

// NETWORK 13
g_AnalogSensor.fbAnalogSensor[E_ASense_Name.TT1004](nSensorID := E_ASense_Name.TT1004, nRawSensor := gIO.ai_EL[1].ch8); // FB_AnalogSensor

// NETWORK 14
g_AnalogSensor.fbAnalogSensor[E_ASense_Name.TT1101](nSensorID := E_ASense_Name.TT1101, nRawSensor := gIO.ai_EL[2].ch3); // FB_AnalogSensor

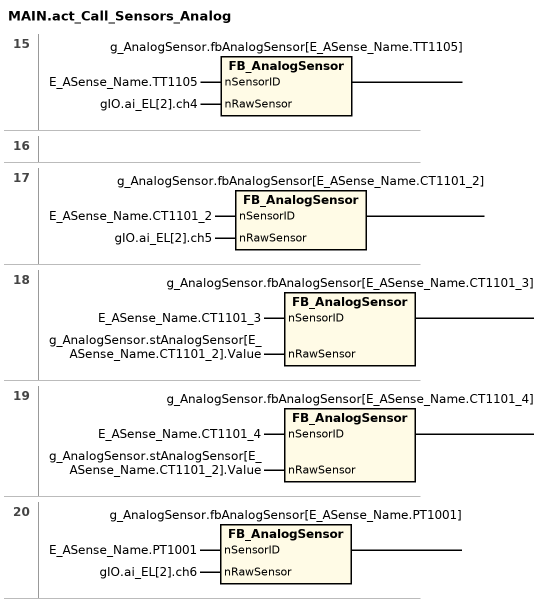
// NETWORK 15
g_AnalogSensor.fbAnalogSensor[E_ASense_Name.TT1105](nSensorID := E_ASense_Name.TT1105, nRawSensor := gIO.ai_EL[2].ch4); // FB_AnalogSensor

// NETWORK 16

// NETWORK 17
g_AnalogSensor.fbAnalogSensor[E_ASense_Name.CT1101_2](nSensorID := E_ASense_Name.CT1101_2, nRawSensor := gIO.ai_EL[2].ch5); // FB_AnalogSensor

// NETWORK 18
g_AnalogSensor.fbAnalogSensor[E_ASense_Name.CT1101_3](nSensorID := E_ASense_Name.CT1101_3, nRawSensor := g_AnalogSensor.stAnalogSensor[E_ASense_Name.CT1101_2].Value); // FB_AnalogSensor

// NETWORK 19
g_AnalogSensor.fbAnalogSensor[E_ASense_Name.CT1101_4](nSensorID := E_ASense_Name.CT1101_4, nRawSensor := g_AnalogSensor.stAnalogSensor[E_ASense_Name.CT1101_2].Value); // FB_AnalogSensor

// NETWORK 20
g_AnalogSensor.fbAnalogSensor[E_ASense_Name.PT1001](nSensorID := E_ASense_Name.PT1001, nRawSensor := gIO.ai_EL[2].ch6); // FB_AnalogSensor
END_ACTION

ACTION act_Call_Sensors_Analog_1:
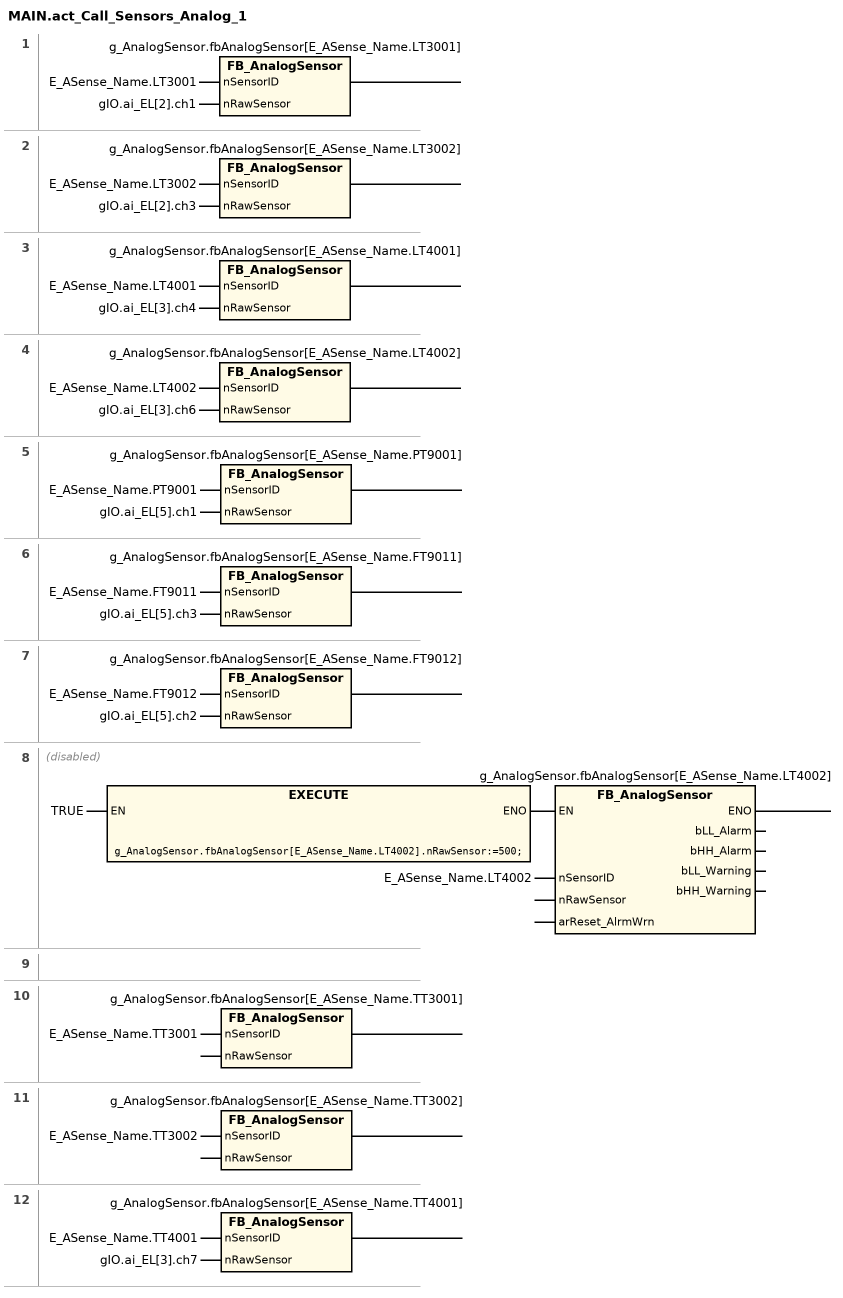
// NETWORK 1
g_AnalogSensor.fbAnalogSensor[E_ASense_Name.LT3001](nSensorID := E_ASense_Name.LT3001, nRawSensor := gIO.ai_EL[2].ch1); // FB_AnalogSensor

// NETWORK 2
g_AnalogSensor.fbAnalogSensor[E_ASense_Name.LT3002](nSensorID := E_ASense_Name.LT3002, nRawSensor := gIO.ai_EL[2].ch3); // FB_AnalogSensor

// NETWORK 3
g_AnalogSensor.fbAnalogSensor[E_ASense_Name.LT4001](nSensorID := E_ASense_Name.LT4001, nRawSensor := gIO.ai_EL[3].ch4); // FB_AnalogSensor

// NETWORK 4
g_AnalogSensor.fbAnalogSensor[E_ASense_Name.LT4002](nSensorID := E_ASense_Name.LT4002, nRawSensor := gIO.ai_EL[3].ch6); // FB_AnalogSensor

// NETWORK 5
g_AnalogSensor.fbAnalogSensor[E_ASense_Name.PT9001](nSensorID := E_ASense_Name.PT9001, nRawSensor := gIO.ai_EL[5].ch1); // FB_AnalogSensor

// NETWORK 6
g_AnalogSensor.fbAnalogSensor[E_ASense_Name.FT9011](nSensorID := E_ASense_Name.FT9011, nRawSensor := gIO.ai_EL[5].ch3); // FB_AnalogSensor

// NETWORK 7
g_AnalogSensor.fbAnalogSensor[E_ASense_Name.FT9012](nSensorID := E_ASense_Name.FT9012, nRawSensor := gIO.ai_EL[5].ch2); // FB_AnalogSensor

// NETWORK 8 (disabled)
// 
// 
// g_AnalogSensor.fbAnalogSensor[E_ASense_Name.LT4002].nRawSensor:=500;
// g_AnalogSensor.fbAnalogSensor[E_ASense_Name.LT4002](nSensorID := E_ASense_Name.LT4002); // FB_AnalogSensor

// NETWORK 9

// NETWORK 10
g_AnalogSensor.fbAnalogSensor[E_ASense_Name.TT3001](nSensorID := E_ASense_Name.TT3001); // FB_AnalogSensor

// NETWORK 11
g_AnalogSensor.fbAnalogSensor[E_ASense_Name.TT3002](nSensorID := E_ASense_Name.TT3002); // FB_AnalogSensor

// NETWORK 12
g_AnalogSensor.fbAnalogSensor[E_ASense_Name.TT4001](nSensorID := E_ASense_Name.TT4001, nRawSensor := gIO.ai_EL[3].ch7); // FB_AnalogSensor

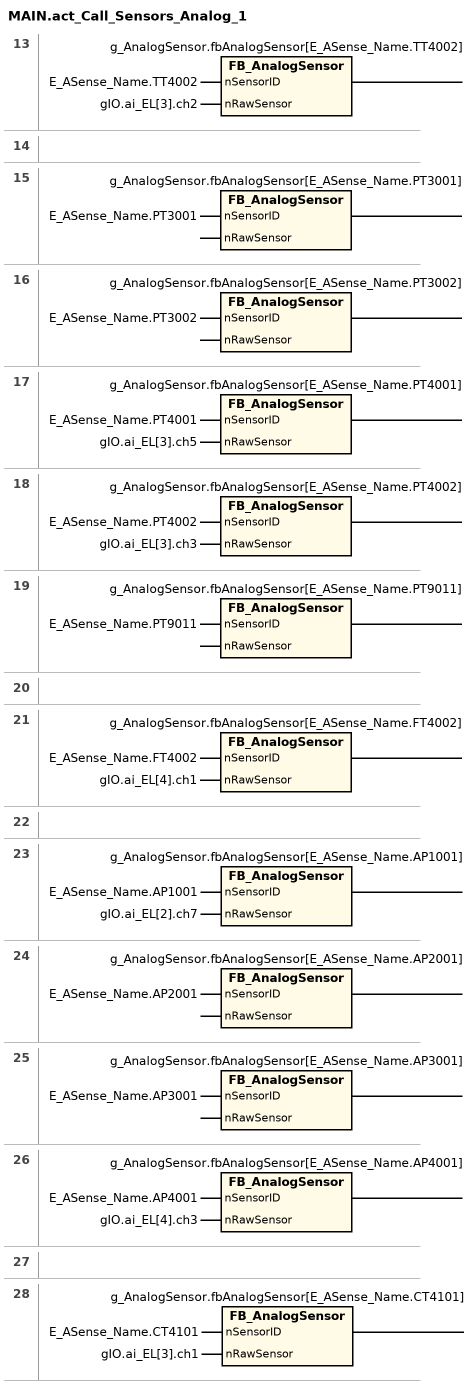
// NETWORK 13
g_AnalogSensor.fbAnalogSensor[E_ASense_Name.TT4002](nSensorID := E_ASense_Name.TT4002, nRawSensor := gIO.ai_EL[3].ch2); // FB_AnalogSensor

// NETWORK 14

// NETWORK 15
g_AnalogSensor.fbAnalogSensor[E_ASense_Name.PT3001](nSensorID := E_ASense_Name.PT3001); // FB_AnalogSensor

// NETWORK 16
g_AnalogSensor.fbAnalogSensor[E_ASense_Name.PT3002](nSensorID := E_ASense_Name.PT3002); // FB_AnalogSensor

// NETWORK 17
g_AnalogSensor.fbAnalogSensor[E_ASense_Name.PT4001](nSensorID := E_ASense_Name.PT4001, nRawSensor := gIO.ai_EL[3].ch5); // FB_AnalogSensor

// NETWORK 18
g_AnalogSensor.fbAnalogSensor[E_ASense_Name.PT4002](nSensorID := E_ASense_Name.PT4002, nRawSensor := gIO.ai_EL[3].ch3); // FB_AnalogSensor

// NETWORK 19
g_AnalogSensor.fbAnalogSensor[E_ASense_Name.PT9011](nSensorID := E_ASense_Name.PT9011); // FB_AnalogSensor

// NETWORK 20

// NETWORK 21
g_AnalogSensor.fbAnalogSensor[E_ASense_Name.FT4002](nSensorID := E_ASense_Name.FT4002, nRawSensor := gIO.ai_EL[4].ch1); // FB_AnalogSensor

// NETWORK 22

// NETWORK 23
g_AnalogSensor.fbAnalogSensor[E_ASense_Name.AP1001](nSensorID := E_ASense_Name.AP1001, nRawSensor := gIO.ai_EL[2].ch7); // FB_AnalogSensor

// NETWORK 24
g_AnalogSensor.fbAnalogSensor[E_ASense_Name.AP2001](nSensorID := E_ASense_Name.AP2001); // FB_AnalogSensor

// NETWORK 25
g_AnalogSensor.fbAnalogSensor[E_ASense_Name.AP3001](nSensorID := E_ASense_Name.AP3001); // FB_AnalogSensor

// NETWORK 26
g_AnalogSensor.fbAnalogSensor[E_ASense_Name.AP4001](nSensorID := E_ASense_Name.AP4001, nRawSensor := gIO.ai_EL[4].ch3); // FB_AnalogSensor

// NETWORK 27

// NETWORK 28
g_AnalogSensor.fbAnalogSensor[E_ASense_Name.CT4101](nSensorID := E_ASense_Name.CT4101, nRawSensor := gIO.ai_EL[3].ch1); // FB_AnalogSensor

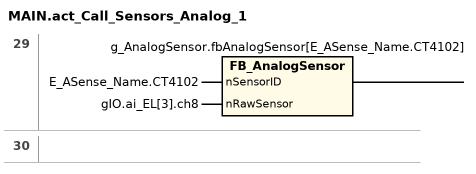
// NETWORK 29
g_AnalogSensor.fbAnalogSensor[E_ASense_Name.CT4102](nSensorID := E_ASense_Name.CT4102, nRawSensor := gIO.ai_EL[3].ch8); // FB_AnalogSensor

// NETWORK 30
END_ACTION

ACTION act_ClientPump_Select:
CASE arCIP_RequestBufer[0].eClient OF
	E_CIP_Usage.eTank_1,
	E_CIP_Usage.eTank_2:;
				eClientPump:=E_Pump_List.P3002;
	E_CIP_Usage.eTank_3,
	E_CIP_Usage.eTank_4:;
				eClientPump:=E_Pump_List.P4002;
	E_CIP_Usage.eLine_Marinada:;
				eClientPump:=E_Pump_List.P3001;
	E_CIP_Usage.eLine_Color:;
				eClientPump:=E_Pump_List.P4001;
	E_CIP_Usage.eTriBlender_Marinada,
	E_CIP_Usage.eTriBlender_Color:;
				eClientPump:=E_Pump_List.TB0001;
	E_CIP_Usage.eLocal:;
				eClientPump:=E_Pump_List.eNotSelected;
END_CASE
END_ACTION

ACTION act_ClientStirrer_Select:
CASE arCIP_RequestBufer[0].eClient OF
	E_CIP_Usage.eTank_1:;
				eClientStirrer:=E_Pump_List.AG3001;
	E_CIP_Usage.eTank_2:;
				eClientStirrer:=E_Pump_List.AG3002;
	E_CIP_Usage.eTank_3:;
				eClientStirrer:=E_Pump_List.AG4001;
	E_CIP_Usage.eTank_4:;
				eClientStirrer:=E_Pump_List.AG4002;
				
	(*E_CIP_Usage.eLine_Marinada:;
	E_CIP_Usage.eLine_Color:;
	E_CIP_Usage.eTriBlender_Marinada,
	E_CIP_Usage.eTriBlender_Color:;*)
ELSE;
	eClientStirrer:=E_Pump_List.eNotSelected;			
END_CASE
END_ACTION

ACTION act_HeatExchenger:
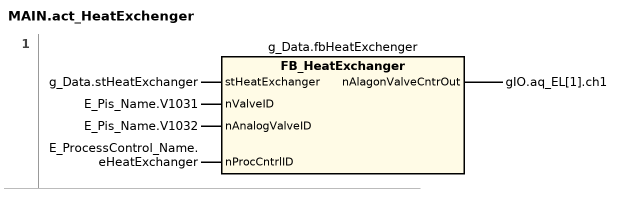
// NETWORK 1
g_Data.fbHeatExchenger(
    stHeatExchanger := g_Data.stHeatExchanger,
    nValveID := E_Pis_Name.V1031,
    nAnalogValveID := E_Pis_Name.V1032,
    nProcCntrlID := E_ProcessControl_Name.eHeatExchanger); // FB_HeatExchanger
gIO.aq_EL[1].ch1 := g_Data.fbHeatExchenger.nAlagonValveCntrOut;
END_ACTION

ACTION act_ResetPumps:
(*ftg_EStop_Fall(CLK:=prg_Safety.ftStateSafe.Q , Q=> );//EStop falling signal
rs_EStopFall(SET:=ftg_EStop_Fall.Q , RESET1:= , Q1=> );
IF rs_EStopFall.Q1 THEN
	FOR nI_1:=1 TO E_Pump_List.last BY 1 DO
		g_Pump.arr_st_Pump[nI_1].bRun_Auto:=FALSE;
	END_FOR
	rs_EStopFall.RESET1:=TRUE;
END_IF
rs_EStopFall.RESET1:=FALSE;*)
;
END_ACTION

ACTION act_Sensors:
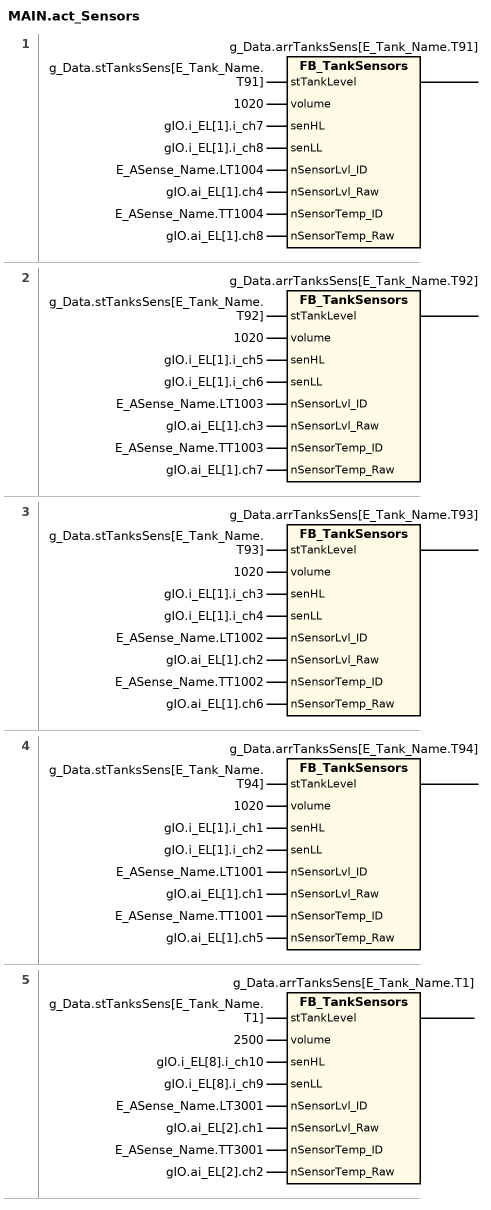
// NETWORK 1
g_Data.arrTanksSens[E_Tank_Name.T91](
    stTankLevel := g_Data.stTanksSens[E_Tank_Name.T91],
    volume := 1020,
    senHL := gIO.i_EL[1].i_ch7,
    senLL := gIO.i_EL[1].i_ch8,
    nSensorLvl_ID := E_ASense_Name.LT1004,
    nSensorLvl_Raw := gIO.ai_EL[1].ch4,
    nSensorTemp_ID := E_ASense_Name.TT1004,
    nSensorTemp_Raw := gIO.ai_EL[1].ch8); // FB_TankSensors

// NETWORK 2
g_Data.arrTanksSens[E_Tank_Name.T92](
    stTankLevel := g_Data.stTanksSens[E_Tank_Name.T92],
    volume := 1020,
    senHL := gIO.i_EL[1].i_ch5,
    senLL := gIO.i_EL[1].i_ch6,
    nSensorLvl_ID := E_ASense_Name.LT1003,
    nSensorLvl_Raw := gIO.ai_EL[1].ch3,
    nSensorTemp_ID := E_ASense_Name.TT1003,
    nSensorTemp_Raw := gIO.ai_EL[1].ch7); // FB_TankSensors

// NETWORK 3
g_Data.arrTanksSens[E_Tank_Name.T93](
    stTankLevel := g_Data.stTanksSens[E_Tank_Name.T93],
    volume := 1020,
    senHL := gIO.i_EL[1].i_ch3,
    senLL := gIO.i_EL[1].i_ch4,
    nSensorLvl_ID := E_ASense_Name.LT1002,
    nSensorLvl_Raw := gIO.ai_EL[1].ch2,
    nSensorTemp_ID := E_ASense_Name.TT1002,
    nSensorTemp_Raw := gIO.ai_EL[1].ch6); // FB_TankSensors

// NETWORK 4
g_Data.arrTanksSens[E_Tank_Name.T94](
    stTankLevel := g_Data.stTanksSens[E_Tank_Name.T94],
    volume := 1020,
    senHL := gIO.i_EL[1].i_ch1,
    senLL := gIO.i_EL[1].i_ch2,
    nSensorLvl_ID := E_ASense_Name.LT1001,
    nSensorLvl_Raw := gIO.ai_EL[1].ch1,
    nSensorTemp_ID := E_ASense_Name.TT1001,
    nSensorTemp_Raw := gIO.ai_EL[1].ch5); // FB_TankSensors

// NETWORK 5
g_Data.arrTanksSens[E_Tank_Name.T1](
    stTankLevel := g_Data.stTanksSens[E_Tank_Name.T1],
    volume := 2500,
    senHL := gIO.i_EL[8].i_ch10,
    senLL := gIO.i_EL[8].i_ch9,
    nSensorLvl_ID := E_ASense_Name.LT3001,
    nSensorLvl_Raw := gIO.ai_EL[2].ch1,
    nSensorTemp_ID := E_ASense_Name.TT3001,
    nSensorTemp_Raw := gIO.ai_EL[2].ch2); // FB_TankSensors

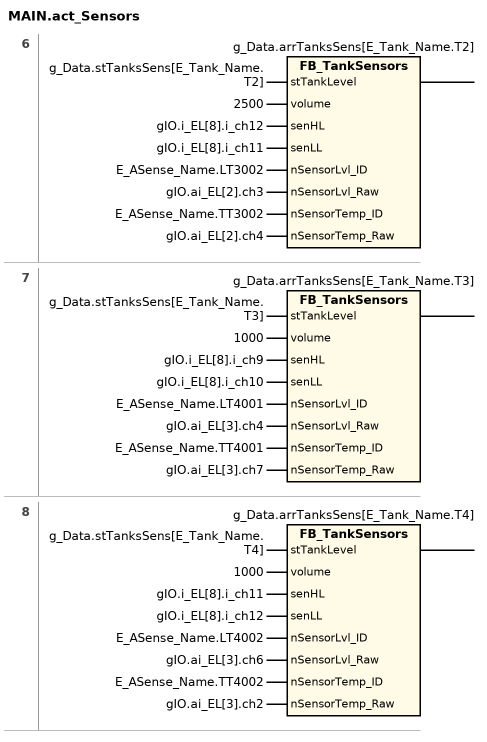
// NETWORK 6
g_Data.arrTanksSens[E_Tank_Name.T2](
    stTankLevel := g_Data.stTanksSens[E_Tank_Name.T2],
    volume := 2500,
    senHL := gIO.i_EL[8].i_ch12,
    senLL := gIO.i_EL[8].i_ch11,
    nSensorLvl_ID := E_ASense_Name.LT3002,
    nSensorLvl_Raw := gIO.ai_EL[2].ch3,
    nSensorTemp_ID := E_ASense_Name.TT3002,
    nSensorTemp_Raw := gIO.ai_EL[2].ch4); // FB_TankSensors

// NETWORK 7
g_Data.arrTanksSens[E_Tank_Name.T3](
    stTankLevel := g_Data.stTanksSens[E_Tank_Name.T3],
    volume := 1000,
    senHL := gIO.i_EL[8].i_ch9,
    senLL := gIO.i_EL[8].i_ch10,
    nSensorLvl_ID := E_ASense_Name.LT4001,
    nSensorLvl_Raw := gIO.ai_EL[3].ch4,
    nSensorTemp_ID := E_ASense_Name.TT4001,
    nSensorTemp_Raw := gIO.ai_EL[3].ch7); // FB_TankSensors

// NETWORK 8
g_Data.arrTanksSens[E_Tank_Name.T4](
    stTankLevel := g_Data.stTanksSens[E_Tank_Name.T4],
    volume := 1000,
    senHL := gIO.i_EL[8].i_ch11,
    senLL := gIO.i_EL[8].i_ch12,
    nSensorLvl_ID := E_ASense_Name.LT4002,
    nSensorLvl_Raw := gIO.ai_EL[3].ch6,
    nSensorTemp_ID := E_ASense_Name.TT4002,
    nSensorTemp_Raw := gIO.ai_EL[3].ch2); // FB_TankSensors
END_ACTION

ACTION act_SetAnalogSens_Test:
//set analog sensors setting only for the test. 
//Later this action should be deleted 
IF NOT bTesting THEN
	//Level
	g_AnalogSensor.stAnalogSensor[E_ASense_Name.LT1004].rawVal_Max:=14350;
	g_AnalogSensor.stAnalogSensor[E_ASense_Name.LT1004].rawVal_Min:=1270;
	g_AnalogSensor.stAnalogSensor[E_ASense_Name.LT1004].outVal_Max:=785;
	g_AnalogSensor.stAnalogSensor[E_ASense_Name.LT1004].outVal_Min:=0;
	g_AnalogSensor.stAnalogSensor[E_ASense_Name.LT1004].outOffset:=73;
	
	g_AnalogSensor.stAnalogSensor[E_ASense_Name.LT1003].rawVal_Max:=14350;
	g_AnalogSensor.stAnalogSensor[E_ASense_Name.LT1003].rawVal_Min:=1270;
	g_AnalogSensor.stAnalogSensor[E_ASense_Name.LT1003].outVal_Max:=785;
	g_AnalogSensor.stAnalogSensor[E_ASense_Name.LT1003].outVal_Min:=0;
	g_AnalogSensor.stAnalogSensor[E_ASense_Name.LT1003].outOffset:=73;
	
	g_AnalogSensor.stAnalogSensor[E_ASense_Name.LT1002].rawVal_Max:=14350;
	g_AnalogSensor.stAnalogSensor[E_ASense_Name.LT1002].rawVal_Min:=1270;
	g_AnalogSensor.stAnalogSensor[E_ASense_Name.LT1002].outVal_Max:=785;
	g_AnalogSensor.stAnalogSensor[E_ASense_Name.LT1002].outVal_Min:=0;
	g_AnalogSensor.stAnalogSensor[E_ASense_Name.LT1002].outOffset:=73;
	
	g_AnalogSensor.stAnalogSensor[E_ASense_Name.LT1001].rawVal_Max:=14350;
	g_AnalogSensor.stAnalogSensor[E_ASense_Name.LT1001].rawVal_Min:=1270;
	g_AnalogSensor.stAnalogSensor[E_ASense_Name.LT1001].outVal_Max:=785;
	g_AnalogSensor.stAnalogSensor[E_ASense_Name.LT1001].outVal_Min:=0;
	g_AnalogSensor.stAnalogSensor[E_ASense_Name.LT1001].outOffset:=73;
	
	//Flow
	g_AnalogSensor.stAnalogSensor[E_ASense_Name.FT1001].rawVal_Max:=10000;
	g_AnalogSensor.stAnalogSensor[E_ASense_Name.FT1001].rawVal_Min:=0;
	g_AnalogSensor.stAnalogSensor[E_ASense_Name.FT1001].outVal_Max:=306;
	g_AnalogSensor.stAnalogSensor[E_ASense_Name.FT1001].outVal_Min:=0;
	g_AnalogSensor.stAnalogSensor[E_ASense_Name.FT1001].outOffset:=0;
	
	g_AnalogSensor.stAnalogSensor[E_ASense_Name.FT1002].rawVal_Max:=10000;
	g_AnalogSensor.stAnalogSensor[E_ASense_Name.FT1002].rawVal_Min:=0;
	g_AnalogSensor.stAnalogSensor[E_ASense_Name.FT1002].outVal_Max:=306;
	g_AnalogSensor.stAnalogSensor[E_ASense_Name.FT1002].outVal_Min:=0;
	g_AnalogSensor.stAnalogSensor[E_ASense_Name.FT1002].outOffset:=0;
	
	////conductivity sensors
	g_AnalogSensor.stAnalogSensor[E_ASense_Name.CT1101].rawVal_Max:=14150;
	g_AnalogSensor.stAnalogSensor[E_ASense_Name.CT1101].rawVal_Min:=305;
	g_AnalogSensor.stAnalogSensor[E_ASense_Name.CT1101].outVal_Max:=14560;
	g_AnalogSensor.stAnalogSensor[E_ASense_Name.CT1101].outVal_Min:=346;
	g_AnalogSensor.stAnalogSensor[E_ASense_Name.CT1101].outOffset:=0;
	(*
	g_AnalogSensor.stAnalogSensor[E_ASense_Name.CT3101].rawVal_Max:=14150;
	g_AnalogSensor.stAnalogSensor[E_ASense_Name.CT3101].rawVal_Min:=305;
	g_AnalogSensor.stAnalogSensor[E_ASense_Name.CT3101].outVal_Max:=14560;
	g_AnalogSensor.stAnalogSensor[E_ASense_Name.CT3101].outVal_Min:=346;
	g_AnalogSensor.stAnalogSensor[E_ASense_Name.CT3101].outOffset:=0;
	*)
	//Temperature sensor
	g_AnalogSensor.stAnalogSensor[E_ASense_Name.TT1001].rawVal_Max:=7470;
	g_AnalogSensor.stAnalogSensor[E_ASense_Name.TT1001].rawVal_Min:=6400;
	g_AnalogSensor.stAnalogSensor[E_ASense_Name.TT1001].outVal_Max:=26;
	g_AnalogSensor.stAnalogSensor[E_ASense_Name.TT1001].outVal_Min:=20.9;
	g_AnalogSensor.stAnalogSensor[E_ASense_Name.TT1001].outOffset:=0;
	
	g_AnalogSensor.stAnalogSensor[E_ASense_Name.TT1002].rawVal_Max:=7470;
	g_AnalogSensor.stAnalogSensor[E_ASense_Name.TT1002].rawVal_Min:=6400;
	g_AnalogSensor.stAnalogSensor[E_ASense_Name.TT1002].outVal_Max:=26;
	g_AnalogSensor.stAnalogSensor[E_ASense_Name.TT1002].outVal_Min:=20.9;
	g_AnalogSensor.stAnalogSensor[E_ASense_Name.TT1002].outOffset:=0;
	
	g_AnalogSensor.stAnalogSensor[E_ASense_Name.TT1003].rawVal_Max:=7470;
	g_AnalogSensor.stAnalogSensor[E_ASense_Name.TT1003].rawVal_Min:=6400;
	g_AnalogSensor.stAnalogSensor[E_ASense_Name.TT1003].outVal_Max:=26;
	g_AnalogSensor.stAnalogSensor[E_ASense_Name.TT1003].outVal_Min:=20.9;
	g_AnalogSensor.stAnalogSensor[E_ASense_Name.TT1003].outOffset:=0;
	
	g_AnalogSensor.stAnalogSensor[E_ASense_Name.TT1004].rawVal_Max:=7470;
	g_AnalogSensor.stAnalogSensor[E_ASense_Name.TT1004].rawVal_Min:=6400;
	g_AnalogSensor.stAnalogSensor[E_ASense_Name.TT1004].outVal_Max:=26;
	g_AnalogSensor.stAnalogSensor[E_ASense_Name.TT1004].outVal_Min:=20.9;
	g_AnalogSensor.stAnalogSensor[E_ASense_Name.TT1004].outOffset:=0;
	
	g_AnalogSensor.stAnalogSensor[E_ASense_Name.TT1101].rawVal_Max:=7470;
	g_AnalogSensor.stAnalogSensor[E_ASense_Name.TT1101].rawVal_Min:=6400;
	g_AnalogSensor.stAnalogSensor[E_ASense_Name.TT1101].outVal_Max:=26;
	g_AnalogSensor.stAnalogSensor[E_ASense_Name.TT1101].outVal_Min:=20.9;
	g_AnalogSensor.stAnalogSensor[E_ASense_Name.TT1101].outOffset:=0;

	bTesting:=TRUE;
END_IF
END_ACTION

ACTION act_SetValves:
//Production tank
	//Tank1
	g_Data.arr_TankValves[1].valOutlet:=	E_Pis_Name.V3016;
	g_Data.arr_TankValves[1].valLine:=		E_Pis_Name.V3017;
	g_Data.arr_TankValves[1].valTriBlender:=E_Pis_Name.V3023;
	g_Data.arr_TankValves[1].valDrain:=		E_Pis_Name.V3024;
	g_Data.arr_TankValves[1].valCIP:=		E_Pis_Name.V3025;
	
	g_Data.arr_LineSourceValves[1].valTankA:=			E_Pis_Name.V3017;
	g_Data.arr_LineSourceValves[1].valTankB:=			E_Pis_Name.V3027;
	g_Data.arr_LineSourceValves[1].valTapWater:=		E_Pis_Name.V_Dummy_LSM_01;
	g_Data.arr_LineSourceValves[1].valTapWater_Drain:=	E_Pis_Name.V_Dummy_LSM_02;
	g_Data.arr_LineSourceValves[1].valTapWater_esle:=	E_Pis_Name.V_Dummy_LSM_05;
	g_Data.arr_LineSourceValves[1].valDrain:=			E_Pis_Name.V3018;
	g_Data.arr_LineSourceValves[1].valCIP:=				E_Pis_Name.V3019;
	g_Data.arr_LineSourceValves[1].valCIP_Sel:=			E_Pis_Name.V_Dummy_LSM_06;
	g_Data.arr_LineSourceValves[1].valBlockWater:=		E_Pis_Name.V_Dummy_LSM_03;
	g_Data.arr_LineSourceValves[1].valWaterSource:=		E_Pis_Name.V_Dummy_LSM_04;
	g_Data.arr_LineSourceValves[1].valWaterSource_Drain:=		E_Pis_Name.V_Dummy_LSM_07;
	
	g_Data.arr_TriBlenderSourceValves[1].valTankA:=				E_Pis_Name.V3023;
	g_Data.arr_TriBlenderSourceValves[1].valTankB:=				E_Pis_Name.V3028;
	g_Data.arr_TriBlenderSourceValves[1].valTapWater:=			E_Pis_Name.V_Dummy_TSM_01;
	g_Data.arr_TriBlenderSourceValves[1].valTapWater_Drain:=	E_Pis_Name.V_Dummy_TSM_02;
	g_Data.arr_TriBlenderSourceValves[1].valTapWater_esle:=		E_Pis_Name.V_Dummy_TSM_03;
	g_Data.arr_TriBlenderSourceValves[1].valDrain:=				E_Pis_Name.V3021;
	g_Data.arr_TriBlenderSourceValves[1].valCIP:=				E_Pis_Name.V3022;
	g_Data.arr_TriBlenderSourceValves[1].valCIP_Sel:=			E_Pis_Name.V3020;
	g_Data.arr_TriBlenderSourceValves[1].valBlockWater:=		E_Pis_Name.V3014;
	g_Data.arr_TriBlenderSourceValves[1].valWaterSource:=		E_Pis_Name.V3113;
	g_Data.arr_TriBlenderSourceValves[1].valWaterSource_Drain:=	E_Pis_Name.V2211;
	
	g_Data.arr_LineTargetValves[1].valTankA:=			E_Pis_Name.V_Dummy_01;//0;
	g_Data.arr_LineTargetValves[1].valTankB:=			E_Pis_Name.V_Dummy_02;//0;
	g_Data.arr_LineTargetValves[1].valDrain:=			E_Pis_Name.V_Dummy_03;//0;
	g_Data.arr_LineTargetValves[1].valCIP:=				E_Pis_Name.V_Dummy_04;//0;
	g_Data.arr_LineTargetValves[1].valTankA_Pipe:=		E_Pis_Name.V_Dummy_05;//0;
	g_Data.arr_LineTargetValves[1].valTankB_Pipe:=		E_Pis_Name.V_Dummy_06;//0;
	
	g_Data.arr_fbTriBlenderTargetValves[1].valTankA:=	E_Pis_Name.V3004;
	g_Data.arr_fbTriBlenderTargetValves[1].valTankB:=	E_Pis_Name.V3010;
	g_Data.arr_fbTriBlenderTargetValves[1].valDrain:=	E_Pis_Name.V3008;
	g_Data.arr_fbTriBlenderTargetValves[1].valCIP:=		E_Pis_Name.V3009;
	g_Data.arr_fbTriBlenderTargetValves[1].valTankA_Pipe:=		E_Pis_Name.v3041;
	g_Data.arr_fbTriBlenderTargetValves[1].valTankB_Pipe:=		E_Pis_Name.v3040;
	
	//Tank2
	g_Data.arr_TankValves[2].valOutlet:=	E_Pis_Name.V3015;
	g_Data.arr_TankValves[2].valLine:=		E_Pis_Name.V3027;
	g_Data.arr_TankValves[2].valTriBlender:=E_Pis_Name.V3028;
	g_Data.arr_TankValves[2].valDrain:=		E_Pis_Name.V3029;
	g_Data.arr_TankValves[2].valCIP:=		E_Pis_Name.V3030;
	
	g_Data.arr_LineSourceValves[2].valTankA:=			E_Pis_Name.V3017;
	g_Data.arr_LineSourceValves[2].valTankB:=			E_Pis_Name.V3027;
	g_Data.arr_LineSourceValves[2].valTapWater:=		E_Pis_Name.V_Dummy_LSM_01;
	g_Data.arr_LineSourceValves[2].valTapWater_Drain:=	E_Pis_Name.V_Dummy_LSM_02;
	g_Data.arr_LineSourceValves[2].valTapWater_esle:=	E_Pis_Name.V_Dummy_LSM_05;
	g_Data.arr_LineSourceValves[2].valDrain:=			E_Pis_Name.V3018;
	g_Data.arr_LineSourceValves[2].valCIP:=				E_Pis_Name.V3019;
	g_Data.arr_LineSourceValves[2].valCIP_Sel:=			E_Pis_Name.V_Dummy_LSM_06;
	g_Data.arr_LineSourceValves[2].valBlockWater:=		E_Pis_Name.V_Dummy_LSM_03;
	g_Data.arr_LineSourceValves[2].valWaterSource:=		E_Pis_Name.V_Dummy_LSM_04;
	g_Data.arr_LineSourceValves[2].valWaterSource_Drain:=		E_Pis_Name.V_Dummy_LSM_07;
	
	
	g_Data.arr_TriBlenderSourceValves[2].valTankA:=				E_Pis_Name.V3023;
	g_Data.arr_TriBlenderSourceValves[2].valTankB:=				E_Pis_Name.V3028;
	g_Data.arr_TriBlenderSourceValves[2].valTapWater:=			E_Pis_Name.V_Dummy_TSM_01;
	g_Data.arr_TriBlenderSourceValves[2].valTapWater_Drain:=	E_Pis_Name.V_Dummy_TSM_02;
	g_Data.arr_TriBlenderSourceValves[2].valTapWater_esle:=		E_Pis_Name.V_Dummy_TSM_03;
	g_Data.arr_TriBlenderSourceValves[2].valDrain:=				E_Pis_Name.V3021;
	g_Data.arr_TriBlenderSourceValves[2].valCIP:=				E_Pis_Name.V3022;
	g_Data.arr_TriBlenderSourceValves[2].valCIP_Sel:=			E_Pis_Name.V3020;
	g_Data.arr_TriBlenderSourceValves[2].valBlockWater:=		E_Pis_Name.V3014;
	g_Data.arr_TriBlenderSourceValves[2].valWaterSource:=		E_Pis_Name.V3113;
	g_Data.arr_TriBlenderSourceValves[2].valWaterSource_Drain:=	E_Pis_Name.V2211;
	
	g_Data.arr_LineTargetValves[2].valTankA:=			E_Pis_Name.V_Dummy_01;//0;
	g_Data.arr_LineTargetValves[2].valTankB:=			E_Pis_Name.V_Dummy_02;//0;
	g_Data.arr_LineTargetValves[2].valDrain:=			E_Pis_Name.V_Dummy_03;//0;
	g_Data.arr_LineTargetValves[2].valCIP:=				E_Pis_Name.V_Dummy_04;//0;
	g_Data.arr_LineTargetValves[2].valTankA_Pipe:=		E_Pis_Name.V_Dummy_05;//0;
	g_Data.arr_LineTargetValves[2].valTankB_Pipe:=		E_Pis_Name.V_Dummy_06;//0;	
	
	(*
	g_Data.arr_LineTargetValves[2].valTankA:=			E_Pis_Name.V_Dummy_07;//0;
	g_Data.arr_LineTargetValves[2].valTankB:=			E_Pis_Name.V_Dummy_08;//0;
	g_Data.arr_LineTargetValves[2].valDrain:=			E_Pis_Name.V_Dummy_09;//0;
	g_Data.arr_LineTargetValves[2].valCIP:=				E_Pis_Name.V_Dummy_10;//0;
	g_Data.arr_LineTargetValves[2].valTankA_Pipe:=		E_Pis_Name.V_Dummy_11;//0;
	g_Data.arr_LineTargetValves[2].valTankB_Pipe:=		E_Pis_Name.V_Dummy_12;//0;
	*)
	
	g_Data.arr_fbTriBlenderTargetValves[2].valTankA:=			E_Pis_Name.V3004;
	g_Data.arr_fbTriBlenderTargetValves[2].valTankB:=			E_Pis_Name.V3010;
	g_Data.arr_fbTriBlenderTargetValves[2].valDrain:=			E_Pis_Name.V3008;
	g_Data.arr_fbTriBlenderTargetValves[2].valCIP:=				E_Pis_Name.V3009;
	g_Data.arr_fbTriBlenderTargetValves[2].valTankA_Pipe:=		E_Pis_Name.V3041;
	g_Data.arr_fbTriBlenderTargetValves[2].valTankB_Pipe:=		E_Pis_Name.V3040;
	
	//Tank3
	g_Data.arr_TankValves[3].valOutlet:=	E_Pis_Name.V4016;
	g_Data.arr_TankValves[3].valLine:=		E_Pis_Name.V4017;
	g_Data.arr_TankValves[3].valTriBlender:=E_Pis_Name.V4023;
	g_Data.arr_TankValves[3].valDrain:=		E_Pis_Name.V4024;
	g_Data.arr_TankValves[3].valCIP:=		E_Pis_Name.V4025;
	
	g_Data.arr_LineSourceValves[3].valTankA:=			E_Pis_Name.V4017;
	g_Data.arr_LineSourceValves[3].valTankB:=			E_Pis_Name.V4027;
	g_Data.arr_LineSourceValves[3].valTapWater:=		E_Pis_Name.V2115;
	g_Data.arr_LineSourceValves[3].valTapWater_Drain:=	E_Pis_Name.V2117;
	g_Data.arr_LineSourceValves[3].valTapWater_esle:=	E_Pis_Name.V2116;
	g_Data.arr_LineSourceValves[3].valDrain:=			E_Pis_Name.V4018;
	g_Data.arr_LineSourceValves[3].valCIP:=				E_Pis_Name.V4019;
	g_Data.arr_LineSourceValves[3].valCIP_Sel:=			E_Pis_Name.V_Dummy_LSC_01;
	g_Data.arr_LineSourceValves[3].valBlockWater:=		E_Pis_Name.V_Dummy_LSC_02;
	g_Data.arr_LineSourceValves[3].valWaterSource:=		E_Pis_Name.V_Dummy_LSC_03;
	g_Data.arr_LineSourceValves[3].valWaterSource_Drain:=		E_Pis_Name.V_Dummy_LSC_04;
	
	g_Data.arr_TriBlenderSourceValves[3].valTankA:=				E_Pis_Name.V4023;
	g_Data.arr_TriBlenderSourceValves[3].valTankB:=				E_Pis_Name.V4028;
	g_Data.arr_TriBlenderSourceValves[3].valTapWater:=			E_Pis_Name.V2116;
	g_Data.arr_TriBlenderSourceValves[3].valTapWater_Drain:=	E_Pis_Name.V2117;
	g_Data.arr_TriBlenderSourceValves[3].valTapWater_esle:=		E_Pis_Name.V2115;
	g_Data.arr_TriBlenderSourceValves[3].valDrain:=				E_Pis_Name.V4021;
	g_Data.arr_TriBlenderSourceValves[3].valCIP:=				E_Pis_Name.V4022;
	g_Data.arr_TriBlenderSourceValves[3].valCIP_Sel:=			E_Pis_Name.V4020;
	g_Data.arr_TriBlenderSourceValves[3].valBlockWater:=		E_Pis_Name.V4014;
	g_Data.arr_TriBlenderSourceValves[3].valWaterSource:=		E_Pis_Name.V2114;
	g_Data.arr_TriBlenderSourceValves[3].valWaterSource_Drain:=	E_Pis_Name.V2112;
	
	g_Data.arr_LineTargetValves[3].valTankA:=	E_Pis_Name.V4034;
	g_Data.arr_LineTargetValves[3].valTankB:=	E_Pis_Name.V4033;
	g_Data.arr_LineTargetValves[3].valDrain:=	E_Pis_Name.V4035;
	g_Data.arr_LineTargetValves[3].valCIP:=		E_Pis_Name.V4036;
	g_Data.arr_LineTargetValves[3].valTankA_Pipe:=		E_Pis_Name.V4041;
	g_Data.arr_LineTargetValves[3].valTankB_Pipe:=		E_Pis_Name.V4040;
	
	g_Data.arr_fbTriBlenderTargetValves[3].valTankA:=	E_Pis_Name.V4004;
	g_Data.arr_fbTriBlenderTargetValves[3].valTankB:=	E_Pis_Name.V4010;
	g_Data.arr_fbTriBlenderTargetValves[3].valDrain:=	E_Pis_Name.V4008;
	g_Data.arr_fbTriBlenderTargetValves[3].valCIP:=		E_Pis_Name.V4009;
	g_Data.arr_fbTriBlenderTargetValves[3].valTankA_Pipe:=		E_Pis_Name.V4041;
	g_Data.arr_fbTriBlenderTargetValves[3].valTankB_Pipe:=		E_Pis_Name.V4040;
	
	//Tank4
	g_Data.arr_TankValves[4].valOutlet:=	E_Pis_Name.V4015;
	g_Data.arr_TankValves[4].valLine:=		E_Pis_Name.V4027;
	g_Data.arr_TankValves[4].valTriBlender:=E_Pis_Name.V4028;
	g_Data.arr_TankValves[4].valDrain:=		E_Pis_Name.V4029;
	g_Data.arr_TankValves[4].valCIP:=		E_Pis_Name.V4030;
	
	g_Data.arr_LineSourceValves[4].valTankA:=			E_Pis_Name.V4017;
	g_Data.arr_LineSourceValves[4].valTankB:=			E_Pis_Name.V4027;
	g_Data.arr_LineSourceValves[4].valTapWater:=		E_Pis_Name.V2115;
	g_Data.arr_LineSourceValves[4].valTapWater_Drain:=	E_Pis_Name.V2117;
	g_Data.arr_LineSourceValves[4].valTapWater_esle:=	E_Pis_Name.V2116;
	g_Data.arr_LineSourceValves[4].valDrain:=			E_Pis_Name.V4018;
	g_Data.arr_LineSourceValves[4].valCIP:=				E_Pis_Name.V4019;
	g_Data.arr_LineSourceValves[4].valCIP_Sel:=			E_Pis_Name.V_Dummy_LSC_01;
	g_Data.arr_LineSourceValves[4].valBlockWater:=		E_Pis_Name.V_Dummy_LSC_02;
	g_Data.arr_LineSourceValves[4].valWaterSource:=		E_Pis_Name.V_Dummy_LSC_03;
	g_Data.arr_LineSourceValves[4].valWaterSource_Drain:=		E_Pis_Name.V_Dummy_LSC_04;
	
	g_Data.arr_TriBlenderSourceValves[4].valTankA:=				E_Pis_Name.V4023;
	g_Data.arr_TriBlenderSourceValves[4].valTankB:=				E_Pis_Name.V4028;
	g_Data.arr_TriBlenderSourceValves[4].valTapWater:=			E_Pis_Name.V2116;
	g_Data.arr_TriBlenderSourceValves[4].valTapWater_Drain:=	E_Pis_Name.V2117;
	g_Data.arr_TriBlenderSourceValves[4].valTapWater_esle:=		E_Pis_Name.V2115;
	g_Data.arr_TriBlenderSourceValves[4].valDrain:=				E_Pis_Name.V4021;
	g_Data.arr_TriBlenderSourceValves[4].valCIP:=				E_Pis_Name.V4022;
	g_Data.arr_TriBlenderSourceValves[4].valCIP_Sel:=			E_Pis_Name.V4020;
	g_Data.arr_TriBlenderSourceValves[4].valBlockWater:=		E_Pis_Name.V4014;
	g_Data.arr_TriBlenderSourceValves[4].valWaterSource:=		E_Pis_Name.V2114;
	g_Data.arr_TriBlenderSourceValves[4].valWaterSource_Drain:=	E_Pis_Name.V2112;
	
	g_Data.arr_LineTargetValves[4].valTankA:=	E_Pis_Name.V4034;
	g_Data.arr_LineTargetValves[4].valTankB:=	E_Pis_Name.V4033;
	g_Data.arr_LineTargetValves[4].valDrain:=	E_Pis_Name.V4035;
	g_Data.arr_LineTargetValves[4].valCIP:=		E_Pis_Name.V4036;
	g_Data.arr_LineTargetValves[4].valTankA_Pipe:=		E_Pis_Name.V4041;
	g_Data.arr_LineTargetValves[4].valTankB_Pipe:=		E_Pis_Name.V4040;
	
	g_Data.arr_fbTriBlenderTargetValves[4].valTankA:=	E_Pis_Name.V4004;
	g_Data.arr_fbTriBlenderTargetValves[4].valTankB:=	E_Pis_Name.V4010;
	g_Data.arr_fbTriBlenderTargetValves[4].valDrain:=	E_Pis_Name.V4008;
	g_Data.arr_fbTriBlenderTargetValves[4].valCIP:=		E_Pis_Name.V4009;
	g_Data.arr_fbTriBlenderTargetValves[4].valTankA_Pipe:=		E_Pis_Name.V4041;
	g_Data.arr_fbTriBlenderTargetValves[4].valTankB_Pipe:=		E_Pis_Name.V4040;
END_ACTION

METHOD m_TankConus_Level_Calculation : REAL
VAR_INPUT
	raw: REAL;

END_VAR
VAR
	kConus: REAL:=0.00000002149 ;
END_VAR
IF raw<1230 THEN;
	//m_TankConus_Level_Calculation:=kConus*raw^3;
ELSE;
	m_TankConus_Level_Calculation:=raw;
END_IF
END_METHOD

METHOD mElementList_SetName : BOOL
VAR_INPUT
END_VAR

VAR
	eASense_Name: E_ASense_Name;
	eProcCntrl: E_ProcessControl_Name;
END_VAR
FOR eASense_Name:=0 TO E_ASense_Name.last DO
	arAnalogSensorNameList[eASense_Name]:=TO_STRING(eASense_Name);
END_FOR

FOR eProcCntrl:=0 TO E_ProcessControl_Name.eProcCntrl_Last DO
	arr_ProcCntrl_NameList[eProcCntrl]:=TO_STRING(eProcCntrl);
	g_ProcControl.arr_stProcCntrl[eProcCntrl].idName:=TO_STRING(eProcCntrl);
END_FOR
END_METHOD

END_PROGRAM

(* stored: Version 1.1.0.1, ProductVersion 3.1.4024.15
   POU MAIN: Id {3441d04c-1b6a-45f8-92c9-effbc902d265}, SpecialFunc None
   Action act_Call_CIP: Id {23177538-beef-46ee-b17f-61590a7b02ee}
   Action act_Call_Elements: Id {2c94e7c7-3832-4cfd-b038-f9562ee8f779}
   Action act_Call_Elements_Imp: Id {5de52cdb-2489-41eb-965b-3474bad12cfe}
   Action act_Call_For_HMI: Id {95962895-82ce-49d5-9aef-33bffa18c9fd}
   Action act_Call_ProcessCntrl: Id {2101a6f8-5f32-44b3-875c-cd379d2d685c}
   Action act_Call_Production: Id {79d1bbce-16ed-4247-ba1c-9331ab9baef9}
   Action act_Call_Pump_TB: Id {5db6818d-58b0-4a03-96bf-e73e0f466a45}
   Action act_Call_Pump_TB_0: Id {91a59c1e-3d38-4546-8bd5-40e12db160d2}
   Action act_Call_Pump_TB_C: Id {fc544244-d2e8-4362-9626-1c2ae87200d0}
   Action act_Call_Pump_TB_CIP: Id {c9a45f93-dfa0-46fa-b0d3-ea3846fef660}
   Action act_Call_Pump_TB_M: Id {c598e0be-4667-4a68-a704-30716d13fee6}
   Action act_Call_Pumps: Id {250d1796-6961-486b-9de7-1fb9e6e9ab7d}
   Action act_Call_ScaleFactor: Id {774d29d4-9ded-47dd-863a-e1e521c0ad31}
   Action act_Call_Sensors_Analog: Id {7ffdbc56-05dc-45ee-9e2a-e9c205335a24}
   Action act_Call_Sensors_Analog_1: Id {c3b256f4-619a-4513-b623-368be1d897cc}
   Action act_ClientPump_Select: Id {480df326-8779-4f2c-832e-de232bda0b87}
   Action act_ClientStirrer_Select: Id {05df8c1d-392d-480e-9db6-d6482e017999}
   Action act_HeatExchenger: Id {bf3394df-98fc-4323-89aa-f243bd329b49}
   Action act_ResetPumps: Id {d6d5f25f-7520-4a69-86f1-bc96d10af8f9}
   Action act_Sensors: Id {8d3d0c01-4d42-45d2-a1c2-ec56cd1d1464}
   Action act_SetAnalogSens_Test: Id {455abcb0-c90c-4f45-9ea9-f7b3ab53cef4}
   Action act_SetValves: Id {606bb271-252e-407f-8120-3b3f040d1b23}
   Method m_TankConus_Level_Calculation: Id {a2410655-ac45-4982-beae-77afb1d1db8e}
   Method mElementList_SetName: Id {fee97784-09c9-4c65-955f-9f389d44d720} *)
